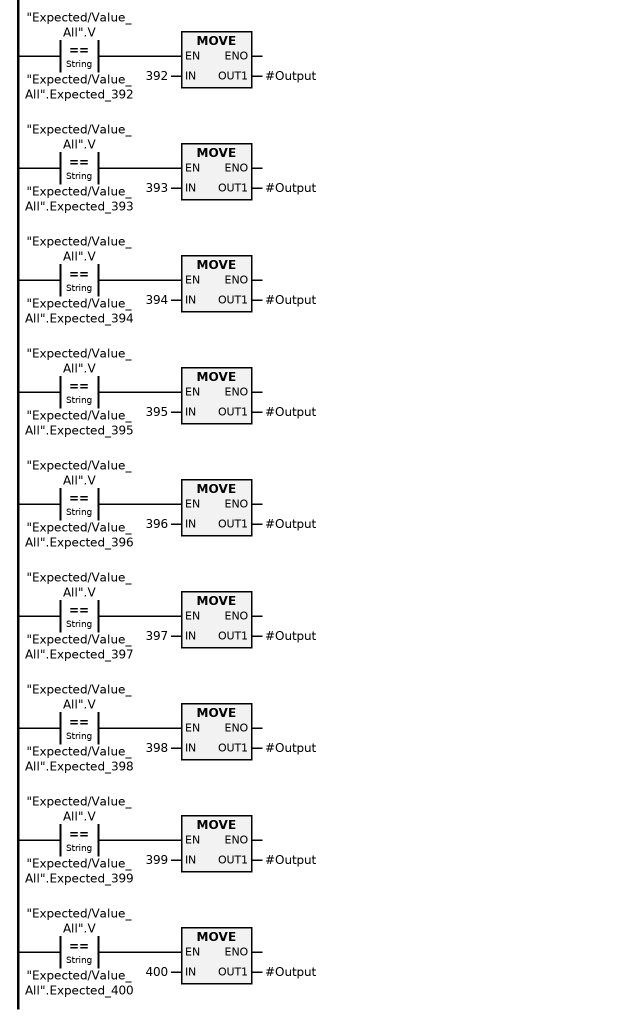
   RUNG wire#powerrail
      { S7_Templates := "SrcType := String" } EQ_Contact(in1 := "Expected/Value_All".V, in2 := "Expected/Value_All".Expected_381)
      Move(in := 381, out1 => #Output)
   END_RUNG
   RUNG wire#powerrail
      { S7_Templates := "SrcType := String" } EQ_Contact(in1 := "Expected/Value_All".V, in2 := "Expected/Value_All".Expected_382)
      Move(in := 382, out1 => #Output)
   END_RUNG
   RUNG wire#powerrail
      { S7_Templates := "SrcType := String" } EQ_Contact(in1 := "Expected/Value_All".V, in2 := "Expected/Value_All".Expected_383)
      Move(in := 383, out1 => #Output)
   END_RUNG
   RUNG wire#powerrail
      { S7_Templates := "SrcType := String" } EQ_Contact(in1 := "Expected/Value_All".V, in2 := "Expected/Value_All".Expected_384)
      Move(in := 384, out1 => #Output)
   END_RUNG
   RUNG wire#powerrail
      { S7_Templates := "SrcType := String" } EQ_Contact(in1 := "Expected/Value_All".V, in2 := "Expected/Value_All".Expected_385)
      Move(in := 385, out1 => #Output)
   END_RUNG
   RUNG wire#powerrail
      { S7_Templates := "SrcType := String" } EQ_Contact(in1 := "Expected/Value_All".V, in2 := "Expected/Value_All".Expected_386)
      Move(in := 386, out1 => #Output)
   END_RUNG
   RUNG wire#powerrail
      { S7_Templates := "SrcType := String" } EQ_Contact(in1 := "Expected/Value_All".V, in2 := "Expected/Value_All".Expected_387)
      Move(in := 387, out1 => #Output)
   END_RUNG
   RUNG wire#powerrail
      { S7_Templates := "SrcType := String" } EQ_Contact(in1 := "Expected/Value_All".V, in2 := "Expected/Value_All".Expected_388)
      Move(in := 388, out1 => #Output)
   END_RUNG
   RUNG wire#powerrail
      { S7_Templates := "SrcType := String" } EQ_Contact(in1 := "Expected/Value_All".V, in2 := "Expected/Value_All".Expected_389)
      Move(in := 389, out1 => #Output)
   END_RUNG
   RUNG wire#powerrail
      { S7_Templates := "SrcType := String" } EQ_Contact(in1 := "Expected/Value_All".V, in2 := "Expected/Value_All".Expected_390)
      Move(in := 390, out1 => #Output)
   END_RUNG
   RUNG wire#powerrail
      { S7_Templates := "SrcType := String" } EQ_Contact(in1 := "Expected/Value_All".V, in2 := "Expected/Value_All".Expected_391)
      Move(in := 391, out1 => #Output)
   END_RUNG
   RUNG wire#powerrail
      { S7_Templates := "SrcType := String" } EQ_Contact(in1 := "Expected/Value_All".V, in2 := "Expected/Value_All".Expected_392)
      Move(in := 392, out1 => #Output)
   END_RUNG
   RUNG wire#powerrail
      { S7_Templates := "SrcType := String" } EQ_Contact(in1 := "Expected/Value_All".V, in2 := "Expected/Value_All".Expected_393)
      Move(in := 393, out1 => #Output)
   END_RUNG
   RUNG wire#powerrail
      { S7_Templates := "SrcType := String" } EQ_Contact(in1 := "Expected/Value_All".V, in2 := "Expected/Value_All".Expected_394)
      Move(in := 394, out1 => #Output)
   END_RUNG
   RUNG wire#powerrail
      { S7_Templates := "SrcType := String" } EQ_Contact(in1 := "Expected/Value_All".V, in2 := "Expected/Value_All".Expected_395)
      Move(in := 395, out1 => #Output)
   END_RUNG
   RUNG wire#powerrail
      { S7_Templates := "SrcType := String" } EQ_Contact(in1 := "Expected/Value_All".V, in2 := "Expected/Value_All".Expected_396)
      Move(in := 396, out1 => #Output)
   END_RUNG
   RUNG wire#powerrail
      { S7_Templates := "SrcType := String" } EQ_Contact(in1 := "Expected/Value_All".V, in2 := "Expected/Value_All".Expected_397)
      Move(in := 397, out1 => #Output)
   END_RUNG
   RUNG wire#powerrail
      { S7_Templates := "SrcType := String" } EQ_Contact(in1 := "Expected/Value_All".V, in2 := "Expected/Value_All".Expected_398)
      Move(in := 398, out1 => #Output)
   END_RUNG
   RUNG wire#powerrail
      { S7_Templates := "SrcType := String" } EQ_Contact(in1 := "Expected/Value_All".V, in2 := "Expected/Value_All".Expected_399)
      Move(in := 399, out1 => #Output)
   END_RUNG
   RUNG wire#powerrail
      { S7_Templates := "SrcType := String" } EQ_Contact(in1 := "Expected/Value_All".V, in2 := "Expected/Value_All".Expected_400)
      Move(in := 400, out1 => #Output)
   END_RUNG
   // the same network as SCL:
   IF "Expected/Value_All".V = "Expected/Value_All".Expected_381 THEN #Output := 381; END_IF;
   IF "Expected/Value_All".V = "Expected/Value_All".Expected_382 THEN #Output := 382; END_IF;
   IF "Expected/Value_All".V = "Expected/Value_All".Expected_383 THEN #Output := 383; END_IF;
   IF "Expected/Value_All".V = "Expected/Value_All".Expected_384 THEN #Output := 384; END_IF;
   IF "Expected/Value_All".V = "Expected/Value_All".Expected_385 THEN #Output := 385; END_IF;
   IF "Expected/Value_All".V = "Expected/Value_All".Expected_386 THEN #Output := 386; END_IF;
   IF "Expected/Value_All".V = "Expected/Value_All".Expected_387 THEN #Output := 387; END_IF;
   IF "Expected/Value_All".V = "Expected/Value_All".Expected_388 THEN #Output := 388; END_IF;
   IF "Expected/Value_All".V = "Expected/Value_All".Expected_389 THEN #Output := 389; END_IF;
   IF "Expected/Value_All".V = "Expected/Value_All".Expected_390 THEN #Output := 390; END_IF;
   IF "Expected/Value_All".V = "Expected/Value_All".Expected_391 THEN #Output := 391; END_IF;
   IF "Expected/Value_All".V = "Expected/Value_All".Expected_392 THEN #Output := 392; END_IF;
   IF "Expected/Value_All".V = "Expected/Value_All".Expected_393 THEN #Output := 393; END_IF;
   IF "Expected/Value_All".V = "Expected/Value_All".Expected_394 THEN #Output := 394; END_IF;
   IF "Expected/Value_All".V = "Expected/Value_All".Expected_395 THEN #Output := 395; END_IF;
   IF "Expected/Value_All".V = "Expected/Value_All".Expected_396 THEN #Output := 396; END_IF;
   IF "Expected/Value_All".V = "Expected/Value_All".Expected_397 THEN #Output := 397; END_IF;
   IF "Expected/Value_All".V = "Expected/Value_All".Expected_398 THEN #Output := 398; END_IF;
   IF "Expected/Value_All".V = "Expected/Value_All".Expected_399 THEN #Output := 399; END_IF;
   IF "Expected/Value_All".V = "Expected/Value_All".Expected_400 THEN #Output := 400; END_IF;
END_REGION

REGION Network 21
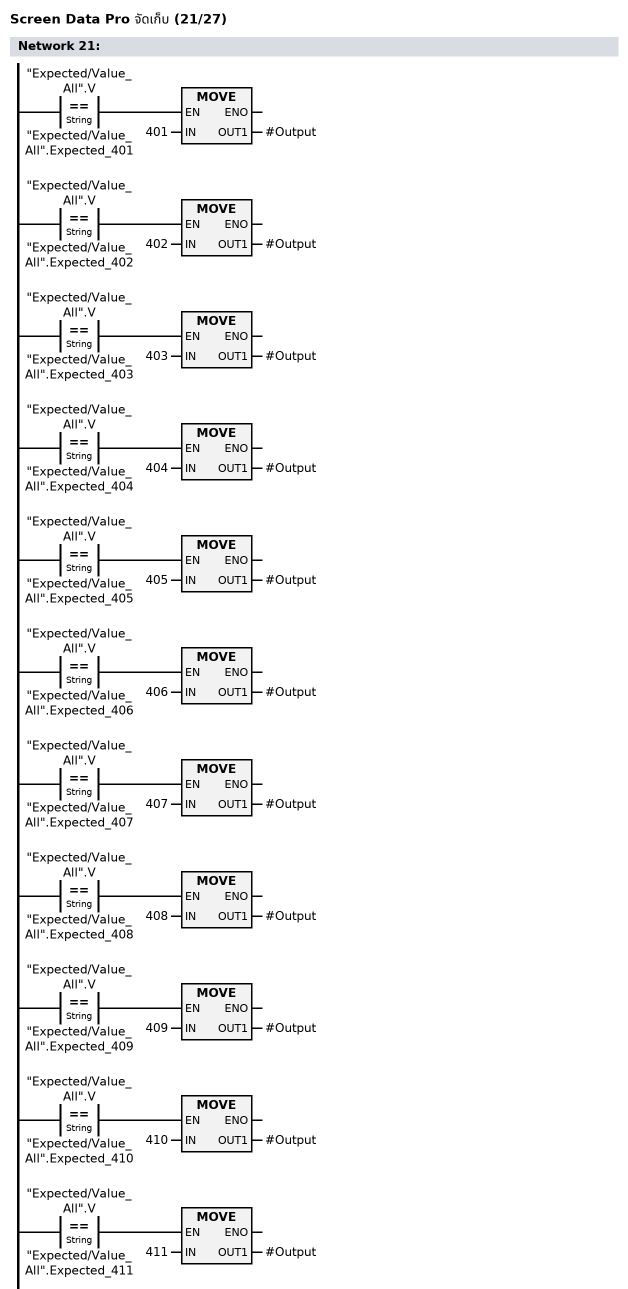
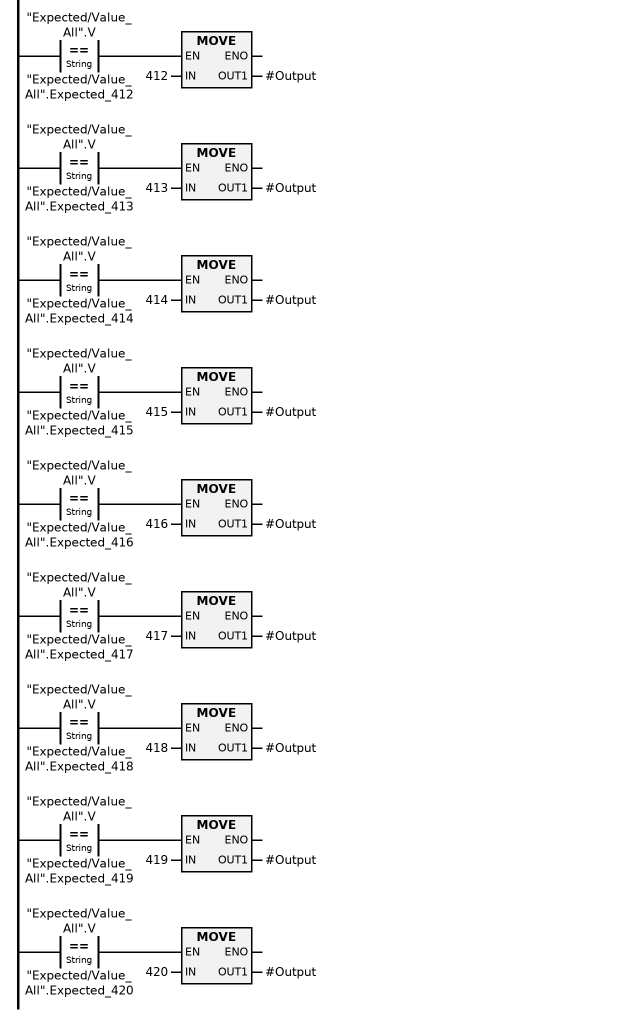
   RUNG wire#powerrail
      { S7_Templates := "SrcType := String" } EQ_Contact(in1 := "Expected/Value_All".V, in2 := "Expected/Value_All".Expected_401)
      Move(in := 401, out1 => #Output)
   END_RUNG
   RUNG wire#powerrail
      { S7_Templates := "SrcType := String" } EQ_Contact(in1 := "Expected/Value_All".V, in2 := "Expected/Value_All".Expected_402)
      Move(in := 402, out1 => #Output)
   END_RUNG
   RUNG wire#powerrail
      { S7_Templates := "SrcType := String" } EQ_Contact(in1 := "Expected/Value_All".V, in2 := "Expected/Value_All".Expected_403)
      Move(in := 403, out1 => #Output)
   END_RUNG
   RUNG wire#powerrail
      { S7_Templates := "SrcType := String" } EQ_Contact(in1 := "Expected/Value_All".V, in2 := "Expected/Value_All".Expected_404)
      Move(in := 404, out1 => #Output)
   END_RUNG
   RUNG wire#powerrail
      { S7_Templates := "SrcType := String" } EQ_Contact(in1 := "Expected/Value_All".V, in2 := "Expected/Value_All".Expected_405)
      Move(in := 405, out1 => #Output)
   END_RUNG
   RUNG wire#powerrail
      { S7_Templates := "SrcType := String" } EQ_Contact(in1 := "Expected/Value_All".V, in2 := "Expected/Value_All".Expected_406)
      Move(in := 406, out1 => #Output)
   END_RUNG
   RUNG wire#powerrail
      { S7_Templates := "SrcType := String" } EQ_Contact(in1 := "Expected/Value_All".V, in2 := "Expected/Value_All".Expected_407)
      Move(in := 407, out1 => #Output)
   END_RUNG
   RUNG wire#powerrail
      { S7_Templates := "SrcType := String" } EQ_Contact(in1 := "Expected/Value_All".V, in2 := "Expected/Value_All".Expected_408)
      Move(in := 408, out1 => #Output)
   END_RUNG
   RUNG wire#powerrail
      { S7_Templates := "SrcType := String" } EQ_Contact(in1 := "Expected/Value_All".V, in2 := "Expected/Value_All".Expected_409)
      Move(in := 409, out1 => #Output)
   END_RUNG
   RUNG wire#powerrail
      { S7_Templates := "SrcType := String" } EQ_Contact(in1 := "Expected/Value_All".V, in2 := "Expected/Value_All".Expected_410)
      Move(in := 410, out1 => #Output)
   END_RUNG
   RUNG wire#powerrail
      { S7_Templates := "SrcType := String" } EQ_Contact(in1 := "Expected/Value_All".V, in2 := "Expected/Value_All".Expected_411)
      Move(in := 411, out1 => #Output)
   END_RUNG
   RUNG wire#powerrail
      { S7_Templates := "SrcType := String" } EQ_Contact(in1 := "Expected/Value_All".V, in2 := "Expected/Value_All".Expected_412)
      Move(in := 412, out1 => #Output)
   END_RUNG
   RUNG wire#powerrail
      { S7_Templates := "SrcType := String" } EQ_Contact(in1 := "Expected/Value_All".V, in2 := "Expected/Value_All".Expected_413)
      Move(in := 413, out1 => #Output)
   END_RUNG
   RUNG wire#powerrail
      { S7_Templates := "SrcType := String" } EQ_Contact(in1 := "Expected/Value_All".V, in2 := "Expected/Value_All".Expected_414)
      Move(in := 414, out1 => #Output)
   END_RUNG
   RUNG wire#powerrail
      { S7_Templates := "SrcType := String" } EQ_Contact(in1 := "Expected/Value_All".V, in2 := "Expected/Value_All".Expected_415)
      Move(in := 415, out1 => #Output)
   END_RUNG
   RUNG wire#powerrail
      { S7_Templates := "SrcType := String" } EQ_Contact(in1 := "Expected/Value_All".V, in2 := "Expected/Value_All".Expected_416)
      Move(in := 416, out1 => #Output)
   END_RUNG
   RUNG wire#powerrail
      { S7_Templates := "SrcType := String" } EQ_Contact(in1 := "Expected/Value_All".V, in2 := "Expected/Value_All".Expected_417)
      Move(in := 417, out1 => #Output)
   END_RUNG
   RUNG wire#powerrail
      { S7_Templates := "SrcType := String" } EQ_Contact(in1 := "Expected/Value_All".V, in2 := "Expected/Value_All".Expected_418)
      Move(in := 418, out1 => #Output)
   END_RUNG
   RUNG wire#powerrail
      { S7_Templates := "SrcType := String" } EQ_Contact(in1 := "Expected/Value_All".V, in2 := "Expected/Value_All".Expected_419)
      Move(in := 419, out1 => #Output)
   END_RUNG
   RUNG wire#powerrail
      { S7_Templates := "SrcType := String" } EQ_Contact(in1 := "Expected/Value_All".V, in2 := "Expected/Value_All".Expected_420)
      Move(in := 420, out1 => #Output)
   END_RUNG
   // the same network as SCL:
   IF "Expected/Value_All".V = "Expected/Value_All".Expected_401 THEN #Output := 401; END_IF;
   IF "Expected/Value_All".V = "Expected/Value_All".Expected_402 THEN #Output := 402; END_IF;
   IF "Expected/Value_All".V = "Expected/Value_All".Expected_403 THEN #Output := 403; END_IF;
   IF "Expected/Value_All".V = "Expected/Value_All".Expected_404 THEN #Output := 404; END_IF;
   IF "Expected/Value_All".V = "Expected/Value_All".Expected_405 THEN #Output := 405; END_IF;
   IF "Expected/Value_All".V = "Expected/Value_All".Expected_406 THEN #Output := 406; END_IF;
   IF "Expected/Value_All".V = "Expected/Value_All".Expected_407 THEN #Output := 407; END_IF;
   IF "Expected/Value_All".V = "Expected/Value_All".Expected_408 THEN #Output := 408; END_IF;
   IF "Expected/Value_All".V = "Expected/Value_All".Expected_409 THEN #Output := 409; END_IF;
   IF "Expected/Value_All".V = "Expected/Value_All".Expected_410 THEN #Output := 410; END_IF;
   IF "Expected/Value_All".V = "Expected/Value_All".Expected_411 THEN #Output := 411; END_IF;
   IF "Expected/Value_All".V = "Expected/Value_All".Expected_412 THEN #Output := 412; END_IF;
   IF "Expected/Value_All".V = "Expected/Value_All".Expected_413 THEN #Output := 413; END_IF;
   IF "Expected/Value_All".V = "Expected/Value_All".Expected_414 THEN #Output := 414; END_IF;
   IF "Expected/Value_All".V = "Expected/Value_All".Expected_415 THEN #Output := 415; END_IF;
   IF "Expected/Value_All".V = "Expected/Value_All".Expected_416 THEN #Output := 416; END_IF;
   IF "Expected/Value_All".V = "Expected/Value_All".Expected_417 THEN #Output := 417; END_IF;
   IF "Expected/Value_All".V = "Expected/Value_All".Expected_418 THEN #Output := 418; END_IF;
   IF "Expected/Value_All".V = "Expected/Value_All".Expected_419 THEN #Output := 419; END_IF;
   IF "Expected/Value_All".V = "Expected/Value_All".Expected_420 THEN #Output := 420; END_IF;
END_REGION

REGION Network 22
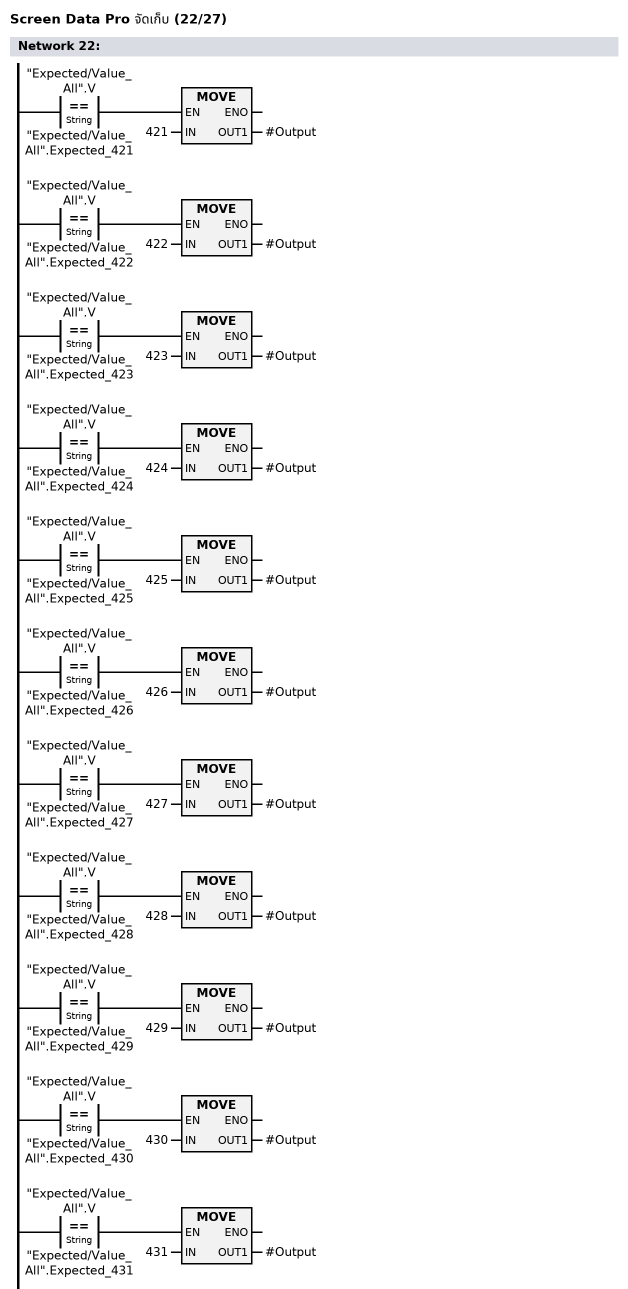
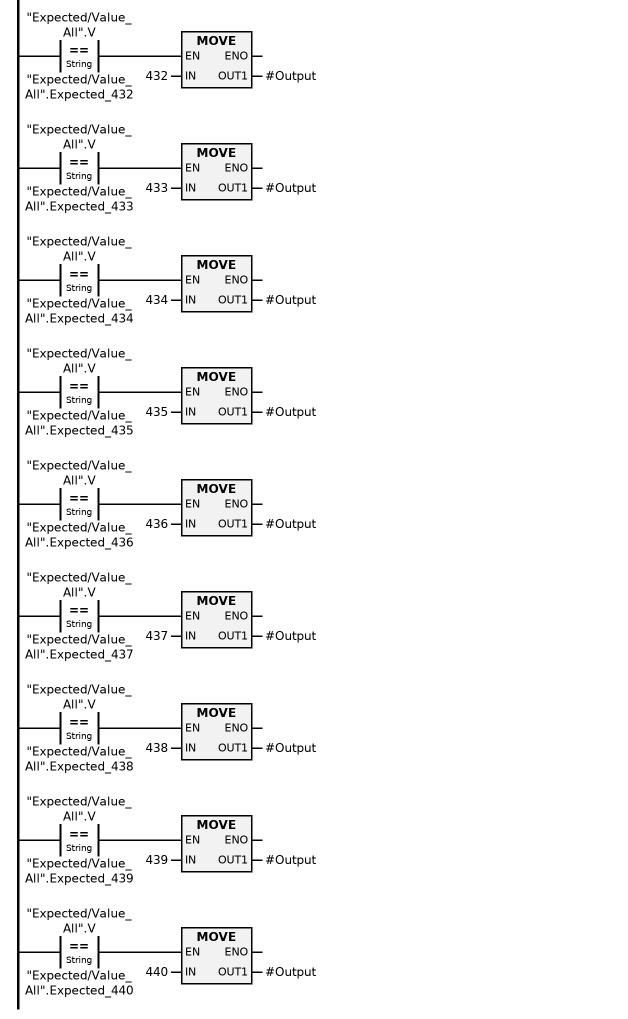
   RUNG wire#powerrail
      { S7_Templates := "SrcType := String" } EQ_Contact(in1 := "Expected/Value_All".V, in2 := "Expected/Value_All".Expected_421)
      Move(in := 421, out1 => #Output)
   END_RUNG
   RUNG wire#powerrail
      { S7_Templates := "SrcType := String" } EQ_Contact(in1 := "Expected/Value_All".V, in2 := "Expected/Value_All".Expected_422)
      Move(in := 422, out1 => #Output)
   END_RUNG
   RUNG wire#powerrail
      { S7_Templates := "SrcType := String" } EQ_Contact(in1 := "Expected/Value_All".V, in2 := "Expected/Value_All".Expected_423)
      Move(in := 423, out1 => #Output)
   END_RUNG
   RUNG wire#powerrail
      { S7_Templates := "SrcType := String" } EQ_Contact(in1 := "Expected/Value_All".V, in2 := "Expected/Value_All".Expected_424)
      Move(in := 424, out1 => #Output)
   END_RUNG
   RUNG wire#powerrail
      { S7_Templates := "SrcType := String" } EQ_Contact(in1 := "Expected/Value_All".V, in2 := "Expected/Value_All".Expected_425)
      Move(in := 425, out1 => #Output)
   END_RUNG
   RUNG wire#powerrail
      { S7_Templates := "SrcType := String" } EQ_Contact(in1 := "Expected/Value_All".V, in2 := "Expected/Value_All".Expected_426)
      Move(in := 426, out1 => #Output)
   END_RUNG
   RUNG wire#powerrail
      { S7_Templates := "SrcType := String" } EQ_Contact(in1 := "Expected/Value_All".V, in2 := "Expected/Value_All".Expected_427)
      Move(in := 427, out1 => #Output)
   END_RUNG
   RUNG wire#powerrail
      { S7_Templates := "SrcType := String" } EQ_Contact(in1 := "Expected/Value_All".V, in2 := "Expected/Value_All".Expected_428)
      Move(in := 428, out1 => #Output)
   END_RUNG
   RUNG wire#powerrail
      { S7_Templates := "SrcType := String" } EQ_Contact(in1 := "Expected/Value_All".V, in2 := "Expected/Value_All".Expected_429)
      Move(in := 429, out1 => #Output)
   END_RUNG
   RUNG wire#powerrail
      { S7_Templates := "SrcType := String" } EQ_Contact(in1 := "Expected/Value_All".V, in2 := "Expected/Value_All".Expected_430)
      Move(in := 430, out1 => #Output)
   END_RUNG
   RUNG wire#powerrail
      { S7_Templates := "SrcType := String" } EQ_Contact(in1 := "Expected/Value_All".V, in2 := "Expected/Value_All".Expected_431)
      Move(in := 431, out1 => #Output)
   END_RUNG
   RUNG wire#powerrail
      { S7_Templates := "SrcType := String" } EQ_Contact(in1 := "Expected/Value_All".V, in2 := "Expected/Value_All".Expected_432)
      Move(in := 432, out1 => #Output)
   END_RUNG
   RUNG wire#powerrail
      { S7_Templates := "SrcType := String" } EQ_Contact(in1 := "Expected/Value_All".V, in2 := "Expected/Value_All".Expected_433)
      Move(in := 433, out1 => #Output)
   END_RUNG
   RUNG wire#powerrail
      { S7_Templates := "SrcType := String" } EQ_Contact(in1 := "Expected/Value_All".V, in2 := "Expected/Value_All".Expected_434)
      Move(in := 434, out1 => #Output)
   END_RUNG
   RUNG wire#powerrail
      { S7_Templates := "SrcType := String" } EQ_Contact(in1 := "Expected/Value_All".V, in2 := "Expected/Value_All".Expected_435)
      Move(in := 435, out1 => #Output)
   END_RUNG
   RUNG wire#powerrail
      { S7_Templates := "SrcType := String" } EQ_Contact(in1 := "Expected/Value_All".V, in2 := "Expected/Value_All".Expected_436)
      Move(in := 436, out1 => #Output)
   END_RUNG
   RUNG wire#powerrail
      { S7_Templates := "SrcType := String" } EQ_Contact(in1 := "Expected/Value_All".V, in2 := "Expected/Value_All".Expected_437)
      Move(in := 437, out1 => #Output)
   END_RUNG
   RUNG wire#powerrail
      { S7_Templates := "SrcType := String" } EQ_Contact(in1 := "Expected/Value_All".V, in2 := "Expected/Value_All".Expected_438)
      Move(in := 438, out1 => #Output)
   END_RUNG
   RUNG wire#powerrail
      { S7_Templates := "SrcType := String" } EQ_Contact(in1 := "Expected/Value_All".V, in2 := "Expected/Value_All".Expected_439)
      Move(in := 439, out1 => #Output)
   END_RUNG
   RUNG wire#powerrail
      { S7_Templates := "SrcType := String" } EQ_Contact(in1 := "Expected/Value_All".V, in2 := "Expected/Value_All".Expected_440)
      Move(in := 440, out1 => #Output)
   END_RUNG
   // the same network as SCL:
   IF "Expected/Value_All".V = "Expected/Value_All".Expected_421 THEN #Output := 421; END_IF;
   IF "Expected/Value_All".V = "Expected/Value_All".Expected_422 THEN #Output := 422; END_IF;
   IF "Expected/Value_All".V = "Expected/Value_All".Expected_423 THEN #Output := 423; END_IF;
   IF "Expected/Value_All".V = "Expected/Value_All".Expected_424 THEN #Output := 424; END_IF;
   IF "Expected/Value_All".V = "Expected/Value_All".Expected_425 THEN #Output := 425; END_IF;
   IF "Expected/Value_All".V = "Expected/Value_All".Expected_426 THEN #Output := 426; END_IF;
   IF "Expected/Value_All".V = "Expected/Value_All".Expected_427 THEN #Output := 427; END_IF;
   IF "Expected/Value_All".V = "Expected/Value_All".Expected_428 THEN #Output := 428; END_IF;
   IF "Expected/Value_All".V = "Expected/Value_All".Expected_429 THEN #Output := 429; END_IF;
   IF "Expected/Value_All".V = "Expected/Value_All".Expected_430 THEN #Output := 430; END_IF;
   IF "Expected/Value_All".V = "Expected/Value_All".Expected_431 THEN #Output := 431; END_IF;
   IF "Expected/Value_All".V = "Expected/Value_All".Expected_432 THEN #Output := 432; END_IF;
   IF "Expected/Value_All".V = "Expected/Value_All".Expected_433 THEN #Output := 433; END_IF;
   IF "Expected/Value_All".V = "Expected/Value_All".Expected_434 THEN #Output := 434; END_IF;
   IF "Expected/Value_All".V = "Expected/Value_All".Expected_435 THEN #Output := 435; END_IF;
   IF "Expected/Value_All".V = "Expected/Value_All".Expected_436 THEN #Output := 436; END_IF;
   IF "Expected/Value_All".V = "Expected/Value_All".Expected_437 THEN #Output := 437; END_IF;
   IF "Expected/Value_All".V = "Expected/Value_All".Expected_438 THEN #Output := 438; END_IF;
   IF "Expected/Value_All".V = "Expected/Value_All".Expected_439 THEN #Output := 439; END_IF;
   IF "Expected/Value_All".V = "Expected/Value_All".Expected_440 THEN #Output := 440; END_IF;
END_REGION

REGION Network 23
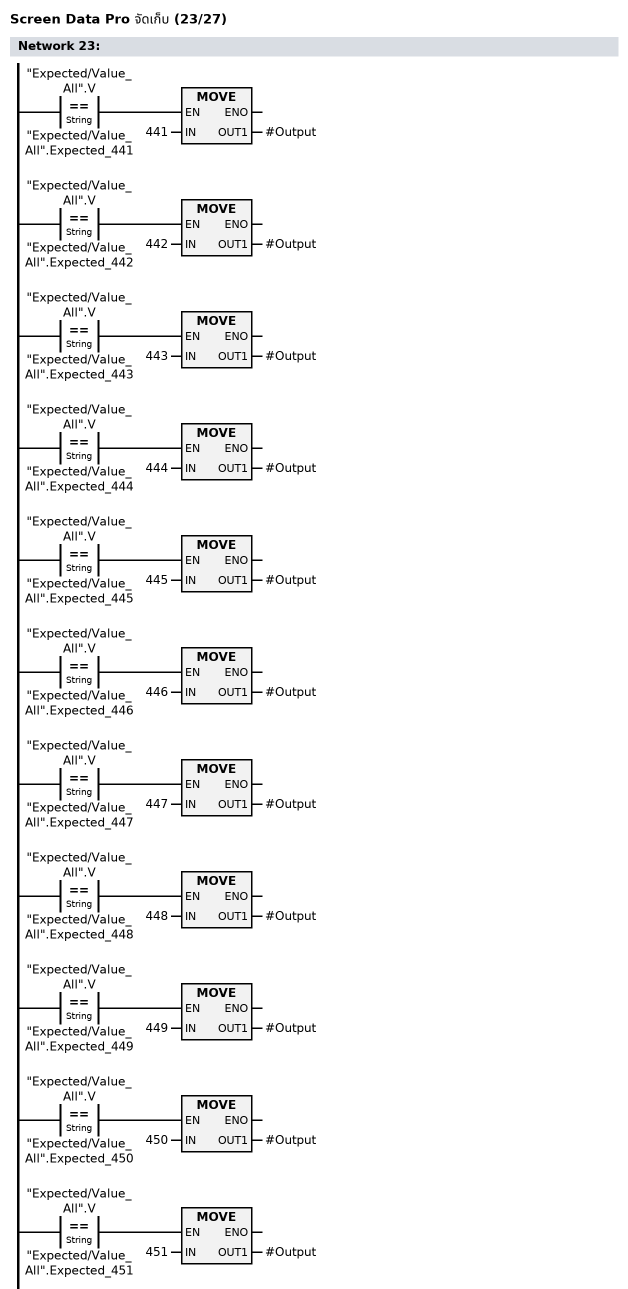
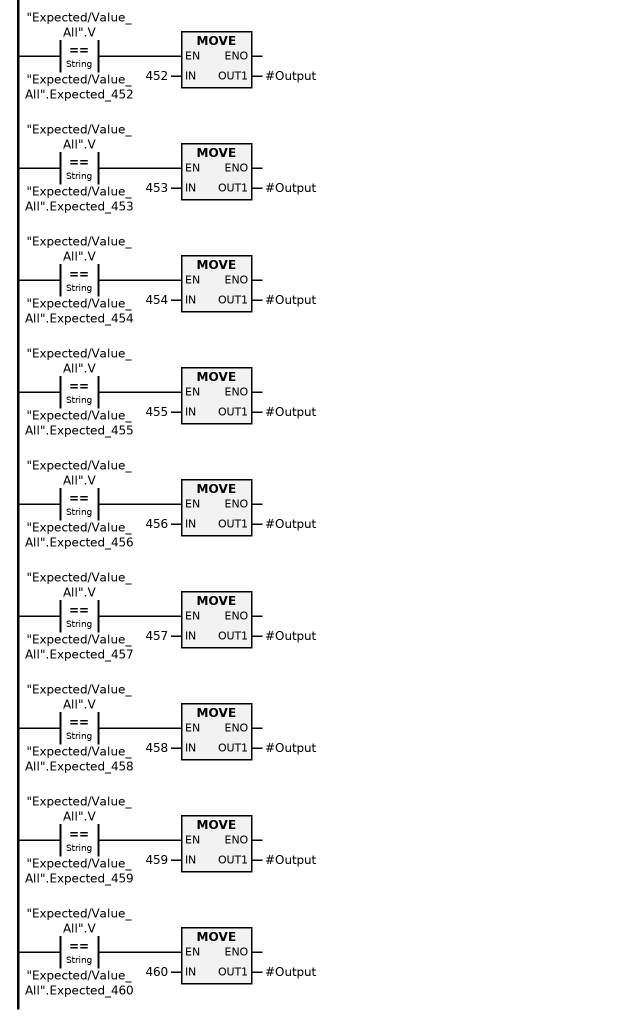
   RUNG wire#powerrail
      { S7_Templates := "SrcType := String" } EQ_Contact(in1 := "Expected/Value_All".V, in2 := "Expected/Value_All".Expected_441)
      Move(in := 441, out1 => #Output)
   END_RUNG
   RUNG wire#powerrail
      { S7_Templates := "SrcType := String" } EQ_Contact(in1 := "Expected/Value_All".V, in2 := "Expected/Value_All".Expected_442)
      Move(in := 442, out1 => #Output)
   END_RUNG
   RUNG wire#powerrail
      { S7_Templates := "SrcType := String" } EQ_Contact(in1 := "Expected/Value_All".V, in2 := "Expected/Value_All".Expected_443)
      Move(in := 443, out1 => #Output)
   END_RUNG
   RUNG wire#powerrail
      { S7_Templates := "SrcType := String" } EQ_Contact(in1 := "Expected/Value_All".V, in2 := "Expected/Value_All".Expected_444)
      Move(in := 444, out1 => #Output)
   END_RUNG
   RUNG wire#powerrail
      { S7_Templates := "SrcType := String" } EQ_Contact(in1 := "Expected/Value_All".V, in2 := "Expected/Value_All".Expected_445)
      Move(in := 445, out1 => #Output)
   END_RUNG
   RUNG wire#powerrail
      { S7_Templates := "SrcType := String" } EQ_Contact(in1 := "Expected/Value_All".V, in2 := "Expected/Value_All".Expected_446)
      Move(in := 446, out1 => #Output)
   END_RUNG
   RUNG wire#powerrail
      { S7_Templates := "SrcType := String" } EQ_Contact(in1 := "Expected/Value_All".V, in2 := "Expected/Value_All".Expected_447)
      Move(in := 447, out1 => #Output)
   END_RUNG
   RUNG wire#powerrail
      { S7_Templates := "SrcType := String" } EQ_Contact(in1 := "Expected/Value_All".V, in2 := "Expected/Value_All".Expected_448)
      Move(in := 448, out1 => #Output)
   END_RUNG
   RUNG wire#powerrail
      { S7_Templates := "SrcType := String" } EQ_Contact(in1 := "Expected/Value_All".V, in2 := "Expected/Value_All".Expected_449)
      Move(in := 449, out1 => #Output)
   END_RUNG
   RUNG wire#powerrail
      { S7_Templates := "SrcType := String" } EQ_Contact(in1 := "Expected/Value_All".V, in2 := "Expected/Value_All".Expected_450)
      Move(in := 450, out1 => #Output)
   END_RUNG
   RUNG wire#powerrail
      { S7_Templates := "SrcType := String" } EQ_Contact(in1 := "Expected/Value_All".V, in2 := "Expected/Value_All".Expected_451)
      Move(in := 451, out1 => #Output)
   END_RUNG
   RUNG wire#powerrail
      { S7_Templates := "SrcType := String" } EQ_Contact(in1 := "Expected/Value_All".V, in2 := "Expected/Value_All".Expected_452)
      Move(in := 452, out1 => #Output)
   END_RUNG
   RUNG wire#powerrail
      { S7_Templates := "SrcType := String" } EQ_Contact(in1 := "Expected/Value_All".V, in2 := "Expected/Value_All".Expected_453)
      Move(in := 453, out1 => #Output)
   END_RUNG
   RUNG wire#powerrail
      { S7_Templates := "SrcType := String" } EQ_Contact(in1 := "Expected/Value_All".V, in2 := "Expected/Value_All".Expected_454)
      Move(in := 454, out1 => #Output)
   END_RUNG
   RUNG wire#powerrail
      { S7_Templates := "SrcType := String" } EQ_Contact(in1 := "Expected/Value_All".V, in2 := "Expected/Value_All".Expected_455)
      Move(in := 455, out1 => #Output)
   END_RUNG
   RUNG wire#powerrail
      { S7_Templates := "SrcType := String" } EQ_Contact(in1 := "Expected/Value_All".V, in2 := "Expected/Value_All".Expected_456)
      Move(in := 456, out1 => #Output)
   END_RUNG
   RUNG wire#powerrail
      { S7_Templates := "SrcType := String" } EQ_Contact(in1 := "Expected/Value_All".V, in2 := "Expected/Value_All".Expected_457)
      Move(in := 457, out1 => #Output)
   END_RUNG
   RUNG wire#powerrail
      { S7_Templates := "SrcType := String" } EQ_Contact(in1 := "Expected/Value_All".V, in2 := "Expected/Value_All".Expected_458)
      Move(in := 458, out1 => #Output)
   END_RUNG
   RUNG wire#powerrail
      { S7_Templates := "SrcType := String" } EQ_Contact(in1 := "Expected/Value_All".V, in2 := "Expected/Value_All".Expected_459)
      Move(in := 459, out1 => #Output)
   END_RUNG
   RUNG wire#powerrail
      { S7_Templates := "SrcType := String" } EQ_Contact(in1 := "Expected/Value_All".V, in2 := "Expected/Value_All".Expected_460)
      Move(in := 460, out1 => #Output)
   END_RUNG
   // the same network as SCL:
   IF "Expected/Value_All".V = "Expected/Value_All".Expected_441 THEN #Output := 441; END_IF;
   IF "Expected/Value_All".V = "Expected/Value_All".Expected_442 THEN #Output := 442; END_IF;
   IF "Expected/Value_All".V = "Expected/Value_All".Expected_443 THEN #Output := 443; END_IF;
   IF "Expected/Value_All".V = "Expected/Value_All".Expected_444 THEN #Output := 444; END_IF;
   IF "Expected/Value_All".V = "Expected/Value_All".Expected_445 THEN #Output := 445; END_IF;
   IF "Expected/Value_All".V = "Expected/Value_All".Expected_446 THEN #Output := 446; END_IF;
   IF "Expected/Value_All".V = "Expected/Value_All".Expected_447 THEN #Output := 447; END_IF;
   IF "Expected/Value_All".V = "Expected/Value_All".Expected_448 THEN #Output := 448; END_IF;
   IF "Expected/Value_All".V = "Expected/Value_All".Expected_449 THEN #Output := 449; END_IF;
   IF "Expected/Value_All".V = "Expected/Value_All".Expected_450 THEN #Output := 450; END_IF;
   IF "Expected/Value_All".V = "Expected/Value_All".Expected_451 THEN #Output := 451; END_IF;
   IF "Expected/Value_All".V = "Expected/Value_All".Expected_452 THEN #Output := 452; END_IF;
   IF "Expected/Value_All".V = "Expected/Value_All".Expected_453 THEN #Output := 453; END_IF;
   IF "Expected/Value_All".V = "Expected/Value_All".Expected_454 THEN #Output := 454; END_IF;
   IF "Expected/Value_All".V = "Expected/Value_All".Expected_455 THEN #Output := 455; END_IF;
   IF "Expected/Value_All".V = "Expected/Value_All".Expected_456 THEN #Output := 456; END_IF;
   IF "Expected/Value_All".V = "Expected/Value_All".Expected_457 THEN #Output := 457; END_IF;
   IF "Expected/Value_All".V = "Expected/Value_All".Expected_458 THEN #Output := 458; END_IF;
   IF "Expected/Value_All".V = "Expected/Value_All".Expected_459 THEN #Output := 459; END_IF;
   IF "Expected/Value_All".V = "Expected/Value_All".Expected_460 THEN #Output := 460; END_IF;
END_REGION

REGION Network 24
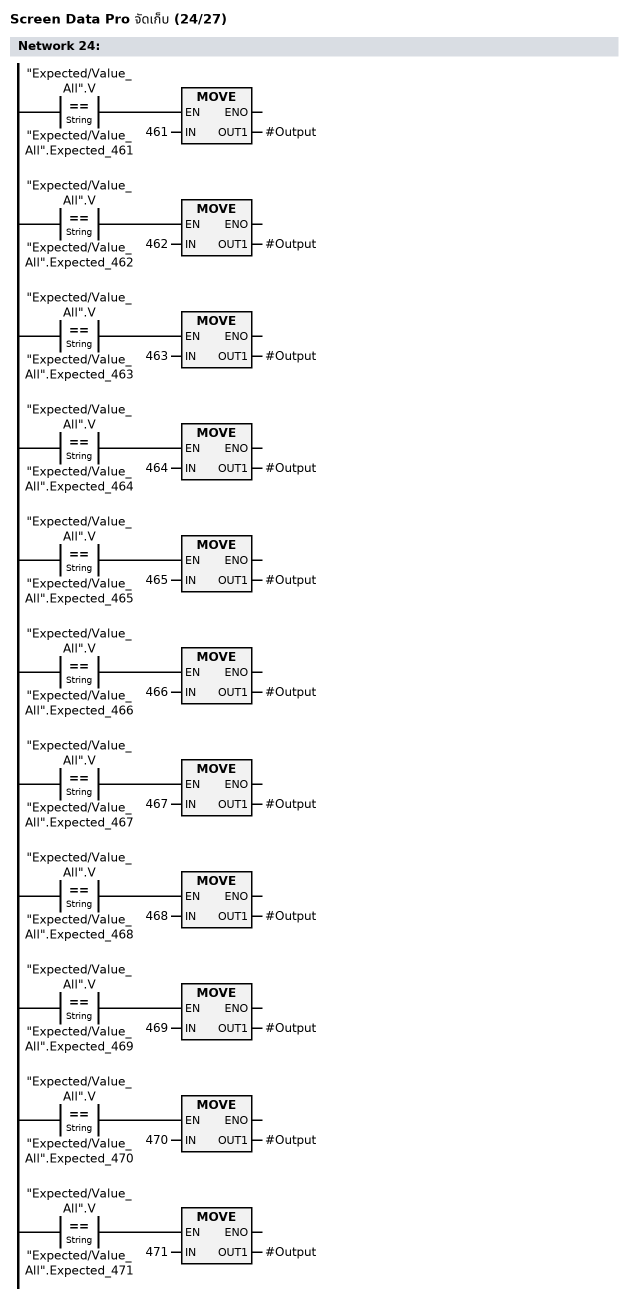
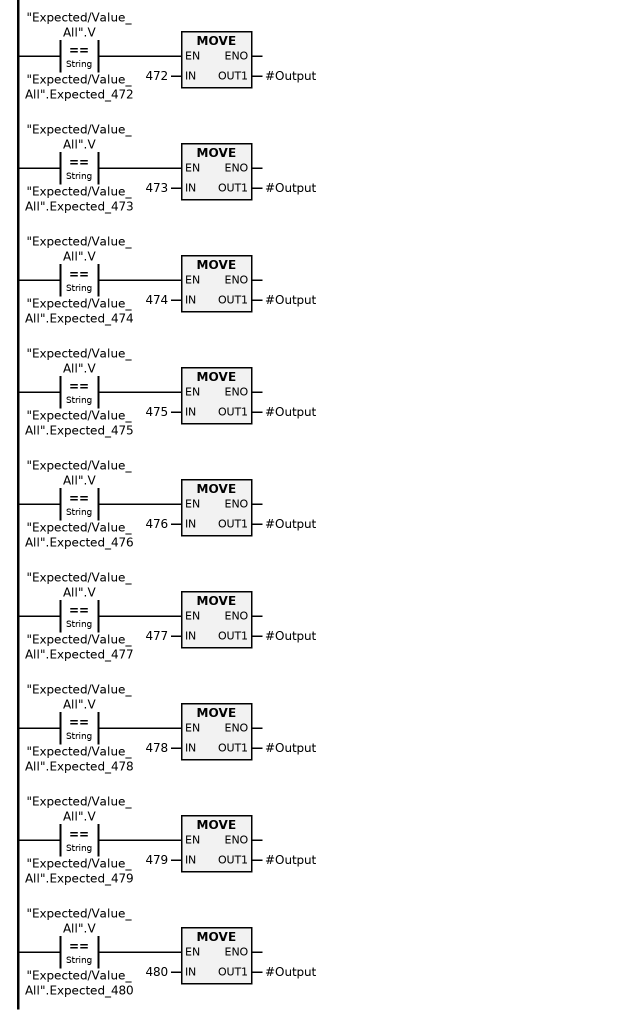
   RUNG wire#powerrail
      { S7_Templates := "SrcType := String" } EQ_Contact(in1 := "Expected/Value_All".V, in2 := "Expected/Value_All".Expected_461)
      Move(in := 461, out1 => #Output)
   END_RUNG
   RUNG wire#powerrail
      { S7_Templates := "SrcType := String" } EQ_Contact(in1 := "Expected/Value_All".V, in2 := "Expected/Value_All".Expected_462)
      Move(in := 462, out1 => #Output)
   END_RUNG
   RUNG wire#powerrail
      { S7_Templates := "SrcType := String" } EQ_Contact(in1 := "Expected/Value_All".V, in2 := "Expected/Value_All".Expected_463)
      Move(in := 463, out1 => #Output)
   END_RUNG
   RUNG wire#powerrail
      { S7_Templates := "SrcType := String" } EQ_Contact(in1 := "Expected/Value_All".V, in2 := "Expected/Value_All".Expected_464)
      Move(in := 464, out1 => #Output)
   END_RUNG
   RUNG wire#powerrail
      { S7_Templates := "SrcType := String" } EQ_Contact(in1 := "Expected/Value_All".V, in2 := "Expected/Value_All".Expected_465)
      Move(in := 465, out1 => #Output)
   END_RUNG
   RUNG wire#powerrail
      { S7_Templates := "SrcType := String" } EQ_Contact(in1 := "Expected/Value_All".V, in2 := "Expected/Value_All".Expected_466)
      Move(in := 466, out1 => #Output)
   END_RUNG
   RUNG wire#powerrail
      { S7_Templates := "SrcType := String" } EQ_Contact(in1 := "Expected/Value_All".V, in2 := "Expected/Value_All".Expected_467)
      Move(in := 467, out1 => #Output)
   END_RUNG
   RUNG wire#powerrail
      { S7_Templates := "SrcType := String" } EQ_Contact(in1 := "Expected/Value_All".V, in2 := "Expected/Value_All".Expected_468)
      Move(in := 468, out1 => #Output)
   END_RUNG
   RUNG wire#powerrail
      { S7_Templates := "SrcType := String" } EQ_Contact(in1 := "Expected/Value_All".V, in2 := "Expected/Value_All".Expected_469)
      Move(in := 469, out1 => #Output)
   END_RUNG
   RUNG wire#powerrail
      { S7_Templates := "SrcType := String" } EQ_Contact(in1 := "Expected/Value_All".V, in2 := "Expected/Value_All".Expected_470)
      Move(in := 470, out1 => #Output)
   END_RUNG
   RUNG wire#powerrail
      { S7_Templates := "SrcType := String" } EQ_Contact(in1 := "Expected/Value_All".V, in2 := "Expected/Value_All".Expected_471)
      Move(in := 471, out1 => #Output)
   END_RUNG
   RUNG wire#powerrail
      { S7_Templates := "SrcType := String" } EQ_Contact(in1 := "Expected/Value_All".V, in2 := "Expected/Value_All".Expected_472)
      Move(in := 472, out1 => #Output)
   END_RUNG
   RUNG wire#powerrail
      { S7_Templates := "SrcType := String" } EQ_Contact(in1 := "Expected/Value_All".V, in2 := "Expected/Value_All".Expected_473)
      Move(in := 473, out1 => #Output)
   END_RUNG
   RUNG wire#powerrail
      { S7_Templates := "SrcType := String" } EQ_Contact(in1 := "Expected/Value_All".V, in2 := "Expected/Value_All".Expected_474)
      Move(in := 474, out1 => #Output)
   END_RUNG
   RUNG wire#powerrail
      { S7_Templates := "SrcType := String" } EQ_Contact(in1 := "Expected/Value_All".V, in2 := "Expected/Value_All".Expected_475)
      Move(in := 475, out1 => #Output)
   END_RUNG
   RUNG wire#powerrail
      { S7_Templates := "SrcType := String" } EQ_Contact(in1 := "Expected/Value_All".V, in2 := "Expected/Value_All".Expected_476)
      Move(in := 476, out1 => #Output)
   END_RUNG
   RUNG wire#powerrail
      { S7_Templates := "SrcType := String" } EQ_Contact(in1 := "Expected/Value_All".V, in2 := "Expected/Value_All".Expected_477)
      Move(in := 477, out1 => #Output)
   END_RUNG
   RUNG wire#powerrail
      { S7_Templates := "SrcType := String" } EQ_Contact(in1 := "Expected/Value_All".V, in2 := "Expected/Value_All".Expected_478)
      Move(in := 478, out1 => #Output)
   END_RUNG
   RUNG wire#powerrail
      { S7_Templates := "SrcType := String" } EQ_Contact(in1 := "Expected/Value_All".V, in2 := "Expected/Value_All".Expected_479)
      Move(in := 479, out1 => #Output)
   END_RUNG
   RUNG wire#powerrail
      { S7_Templates := "SrcType := String" } EQ_Contact(in1 := "Expected/Value_All".V, in2 := "Expected/Value_All".Expected_480)
      Move(in := 480, out1 => #Output)
   END_RUNG
   // the same network as SCL:
   IF "Expected/Value_All".V = "Expected/Value_All".Expected_461 THEN #Output := 461; END_IF;
   IF "Expected/Value_All".V = "Expected/Value_All".Expected_462 THEN #Output := 462; END_IF;
   IF "Expected/Value_All".V = "Expected/Value_All".Expected_463 THEN #Output := 463; END_IF;
   IF "Expected/Value_All".V = "Expected/Value_All".Expected_464 THEN #Output := 464; END_IF;
   IF "Expected/Value_All".V = "Expected/Value_All".Expected_465 THEN #Output := 465; END_IF;
   IF "Expected/Value_All".V = "Expected/Value_All".Expected_466 THEN #Output := 466; END_IF;
   IF "Expected/Value_All".V = "Expected/Value_All".Expected_467 THEN #Output := 467; END_IF;
   IF "Expected/Value_All".V = "Expected/Value_All".Expected_468 THEN #Output := 468; END_IF;
   IF "Expected/Value_All".V = "Expected/Value_All".Expected_469 THEN #Output := 469; END_IF;
   IF "Expected/Value_All".V = "Expected/Value_All".Expected_470 THEN #Output := 470; END_IF;
   IF "Expected/Value_All".V = "Expected/Value_All".Expected_471 THEN #Output := 471; END_IF;
   IF "Expected/Value_All".V = "Expected/Value_All".Expected_472 THEN #Output := 472; END_IF;
   IF "Expected/Value_All".V = "Expected/Value_All".Expected_473 THEN #Output := 473; END_IF;
   IF "Expected/Value_All".V = "Expected/Value_All".Expected_474 THEN #Output := 474; END_IF;
   IF "Expected/Value_All".V = "Expected/Value_All".Expected_475 THEN #Output := 475; END_IF;
   IF "Expected/Value_All".V = "Expected/Value_All".Expected_476 THEN #Output := 476; END_IF;
   IF "Expected/Value_All".V = "Expected/Value_All".Expected_477 THEN #Output := 477; END_IF;
   IF "Expected/Value_All".V = "Expected/Value_All".Expected_478 THEN #Output := 478; END_IF;
   IF "Expected/Value_All".V = "Expected/Value_All".Expected_479 THEN #Output := 479; END_IF;
   IF "Expected/Value_All".V = "Expected/Value_All".Expected_480 THEN #Output := 480; END_IF;
END_REGION

REGION Network 25
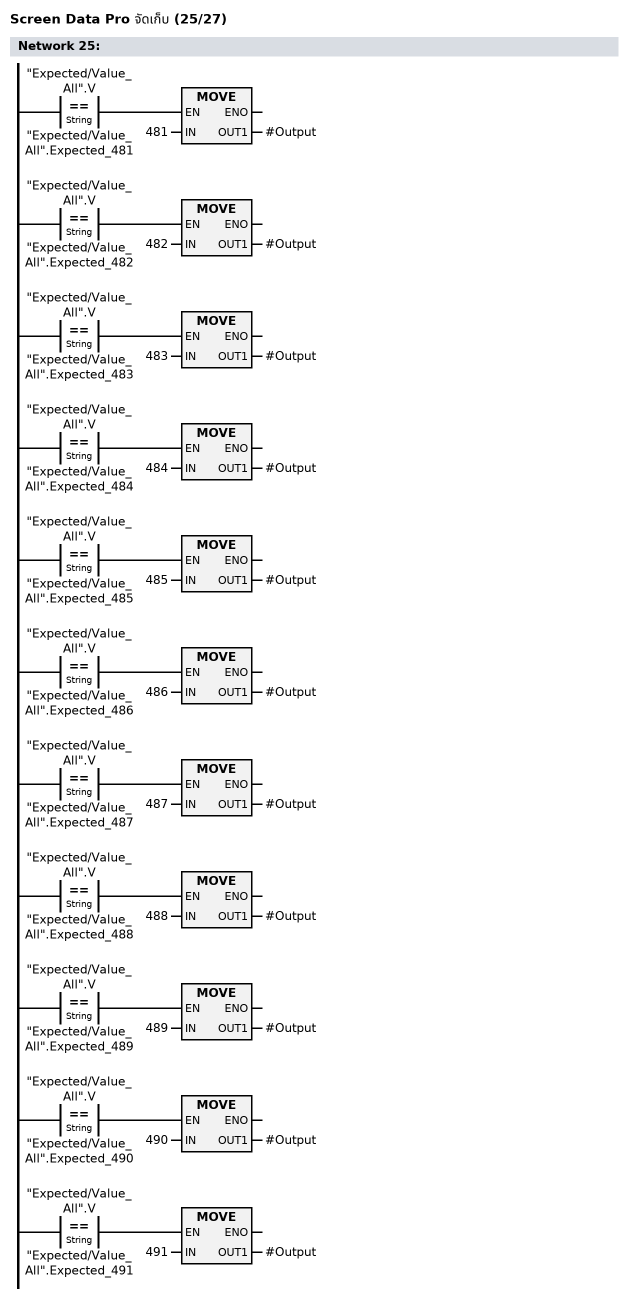
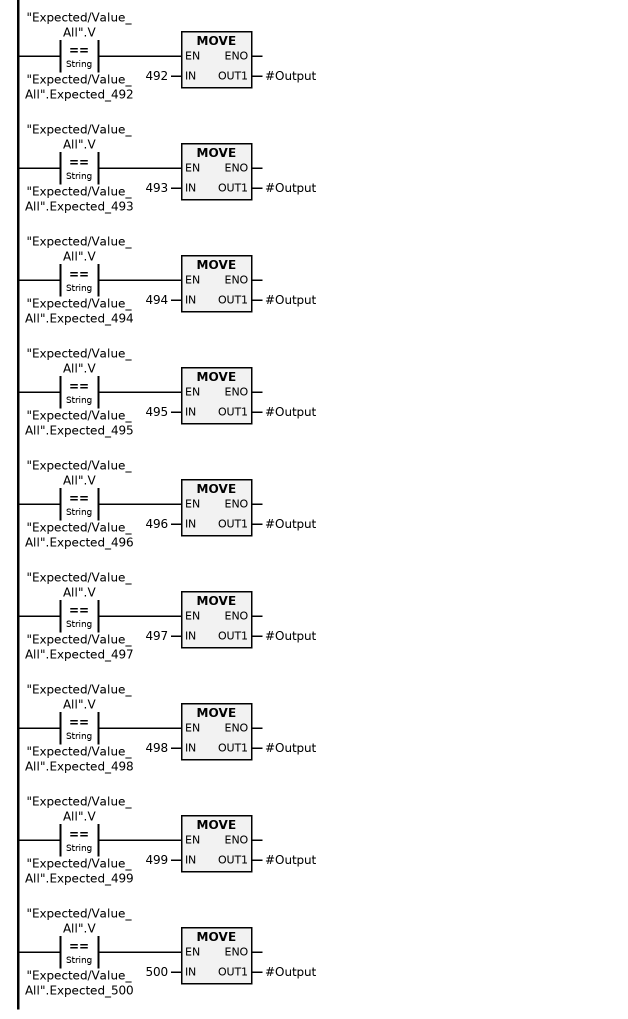
   RUNG wire#powerrail
      { S7_Templates := "SrcType := String" } EQ_Contact(in1 := "Expected/Value_All".V, in2 := "Expected/Value_All".Expected_481)
      Move(in := 481, out1 => #Output)
   END_RUNG
   RUNG wire#powerrail
      { S7_Templates := "SrcType := String" } EQ_Contact(in1 := "Expected/Value_All".V, in2 := "Expected/Value_All".Expected_482)
      Move(in := 482, out1 => #Output)
   END_RUNG
   RUNG wire#powerrail
      { S7_Templates := "SrcType := String" } EQ_Contact(in1 := "Expected/Value_All".V, in2 := "Expected/Value_All".Expected_483)
      Move(in := 483, out1 => #Output)
   END_RUNG
   RUNG wire#powerrail
      { S7_Templates := "SrcType := String" } EQ_Contact(in1 := "Expected/Value_All".V, in2 := "Expected/Value_All".Expected_484)
      Move(in := 484, out1 => #Output)
   END_RUNG
   RUNG wire#powerrail
      { S7_Templates := "SrcType := String" } EQ_Contact(in1 := "Expected/Value_All".V, in2 := "Expected/Value_All".Expected_485)
      Move(in := 485, out1 => #Output)
   END_RUNG
   RUNG wire#powerrail
      { S7_Templates := "SrcType := String" } EQ_Contact(in1 := "Expected/Value_All".V, in2 := "Expected/Value_All".Expected_486)
      Move(in := 486, out1 => #Output)
   END_RUNG
   RUNG wire#powerrail
      { S7_Templates := "SrcType := String" } EQ_Contact(in1 := "Expected/Value_All".V, in2 := "Expected/Value_All".Expected_487)
      Move(in := 487, out1 => #Output)
   END_RUNG
   RUNG wire#powerrail
      { S7_Templates := "SrcType := String" } EQ_Contact(in1 := "Expected/Value_All".V, in2 := "Expected/Value_All".Expected_488)
      Move(in := 488, out1 => #Output)
   END_RUNG
   RUNG wire#powerrail
      { S7_Templates := "SrcType := String" } EQ_Contact(in1 := "Expected/Value_All".V, in2 := "Expected/Value_All".Expected_489)
      Move(in := 489, out1 => #Output)
   END_RUNG
   RUNG wire#powerrail
      { S7_Templates := "SrcType := String" } EQ_Contact(in1 := "Expected/Value_All".V, in2 := "Expected/Value_All".Expected_490)
      Move(in := 490, out1 => #Output)
   END_RUNG
   RUNG wire#powerrail
      { S7_Templates := "SrcType := String" } EQ_Contact(in1 := "Expected/Value_All".V, in2 := "Expected/Value_All".Expected_491)
      Move(in := 491, out1 => #Output)
   END_RUNG
   RUNG wire#powerrail
      { S7_Templates := "SrcType := String" } EQ_Contact(in1 := "Expected/Value_All".V, in2 := "Expected/Value_All".Expected_492)
      Move(in := 492, out1 => #Output)
   END_RUNG
   RUNG wire#powerrail
      { S7_Templates := "SrcType := String" } EQ_Contact(in1 := "Expected/Value_All".V, in2 := "Expected/Value_All".Expected_493)
      Move(in := 493, out1 => #Output)
   END_RUNG
   RUNG wire#powerrail
      { S7_Templates := "SrcType := String" } EQ_Contact(in1 := "Expected/Value_All".V, in2 := "Expected/Value_All".Expected_494)
      Move(in := 494, out1 => #Output)
   END_RUNG
   RUNG wire#powerrail
      { S7_Templates := "SrcType := String" } EQ_Contact(in1 := "Expected/Value_All".V, in2 := "Expected/Value_All".Expected_495)
      Move(in := 495, out1 => #Output)
   END_RUNG
   RUNG wire#powerrail
      { S7_Templates := "SrcType := String" } EQ_Contact(in1 := "Expected/Value_All".V, in2 := "Expected/Value_All".Expected_496)
      Move(in := 496, out1 => #Output)
   END_RUNG
   RUNG wire#powerrail
      { S7_Templates := "SrcType := String" } EQ_Contact(in1 := "Expected/Value_All".V, in2 := "Expected/Value_All".Expected_497)
      Move(in := 497, out1 => #Output)
   END_RUNG
   RUNG wire#powerrail
      { S7_Templates := "SrcType := String" } EQ_Contact(in1 := "Expected/Value_All".V, in2 := "Expected/Value_All".Expected_498)
      Move(in := 498, out1 => #Output)
   END_RUNG
   RUNG wire#powerrail
      { S7_Templates := "SrcType := String" } EQ_Contact(in1 := "Expected/Value_All".V, in2 := "Expected/Value_All".Expected_499)
      Move(in := 499, out1 => #Output)
   END_RUNG
   RUNG wire#powerrail
      { S7_Templates := "SrcType := String" } EQ_Contact(in1 := "Expected/Value_All".V, in2 := "Expected/Value_All".Expected_500)
      Move(in := 500, out1 => #Output)
   END_RUNG
   // the same network as SCL:
   IF "Expected/Value_All".V = "Expected/Value_All".Expected_481 THEN #Output := 481; END_IF;
   IF "Expected/Value_All".V = "Expected/Value_All".Expected_482 THEN #Output := 482; END_IF;
   IF "Expected/Value_All".V = "Expected/Value_All".Expected_483 THEN #Output := 483; END_IF;
   IF "Expected/Value_All".V = "Expected/Value_All".Expected_484 THEN #Output := 484; END_IF;
   IF "Expected/Value_All".V = "Expected/Value_All".Expected_485 THEN #Output := 485; END_IF;
   IF "Expected/Value_All".V = "Expected/Value_All".Expected_486 THEN #Output := 486; END_IF;
   IF "Expected/Value_All".V = "Expected/Value_All".Expected_487 THEN #Output := 487; END_IF;
   IF "Expected/Value_All".V = "Expected/Value_All".Expected_488 THEN #Output := 488; END_IF;
   IF "Expected/Value_All".V = "Expected/Value_All".Expected_489 THEN #Output := 489; END_IF;
   IF "Expected/Value_All".V = "Expected/Value_All".Expected_490 THEN #Output := 490; END_IF;
   IF "Expected/Value_All".V = "Expected/Value_All".Expected_491 THEN #Output := 491; END_IF;
   IF "Expected/Value_All".V = "Expected/Value_All".Expected_492 THEN #Output := 492; END_IF;
   IF "Expected/Value_All".V = "Expected/Value_All".Expected_493 THEN #Output := 493; END_IF;
   IF "Expected/Value_All".V = "Expected/Value_All".Expected_494 THEN #Output := 494; END_IF;
   IF "Expected/Value_All".V = "Expected/Value_All".Expected_495 THEN #Output := 495; END_IF;
   IF "Expected/Value_All".V = "Expected/Value_All".Expected_496 THEN #Output := 496; END_IF;
   IF "Expected/Value_All".V = "Expected/Value_All".Expected_497 THEN #Output := 497; END_IF;
   IF "Expected/Value_All".V = "Expected/Value_All".Expected_498 THEN #Output := 498; END_IF;
   IF "Expected/Value_All".V = "Expected/Value_All".Expected_499 THEN #Output := 499; END_IF;
   IF "Expected/Value_All".V = "Expected/Value_All".Expected_500 THEN #Output := 500; END_IF;
END_REGION

REGION Network 26
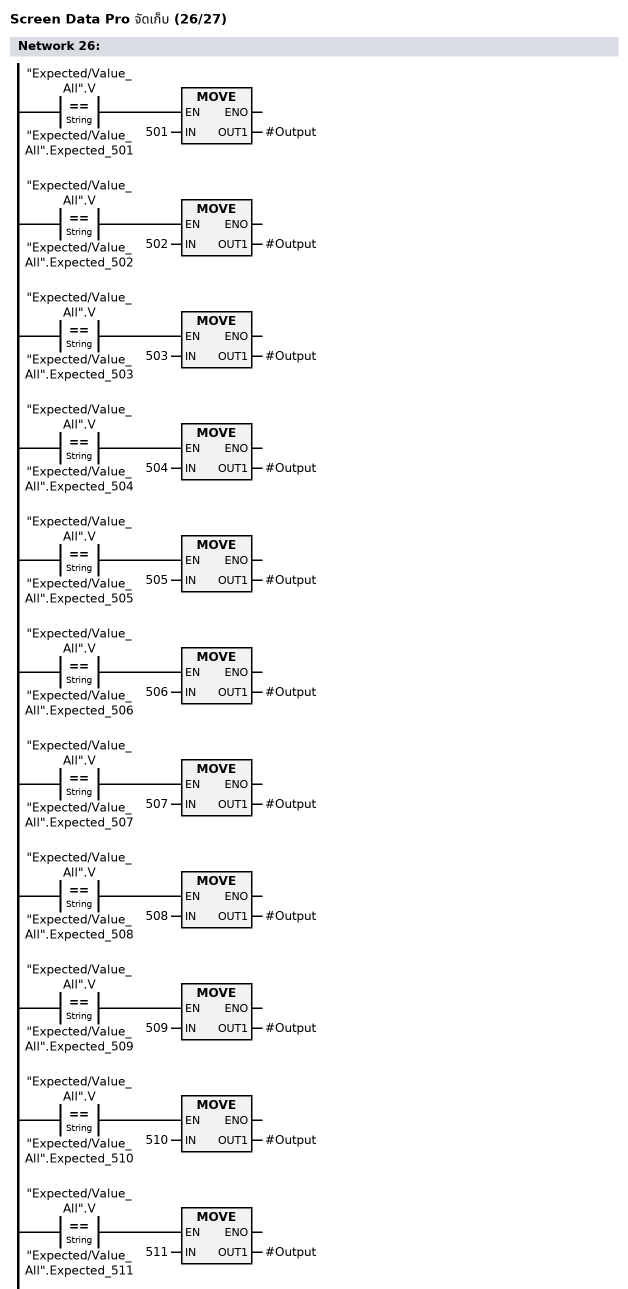
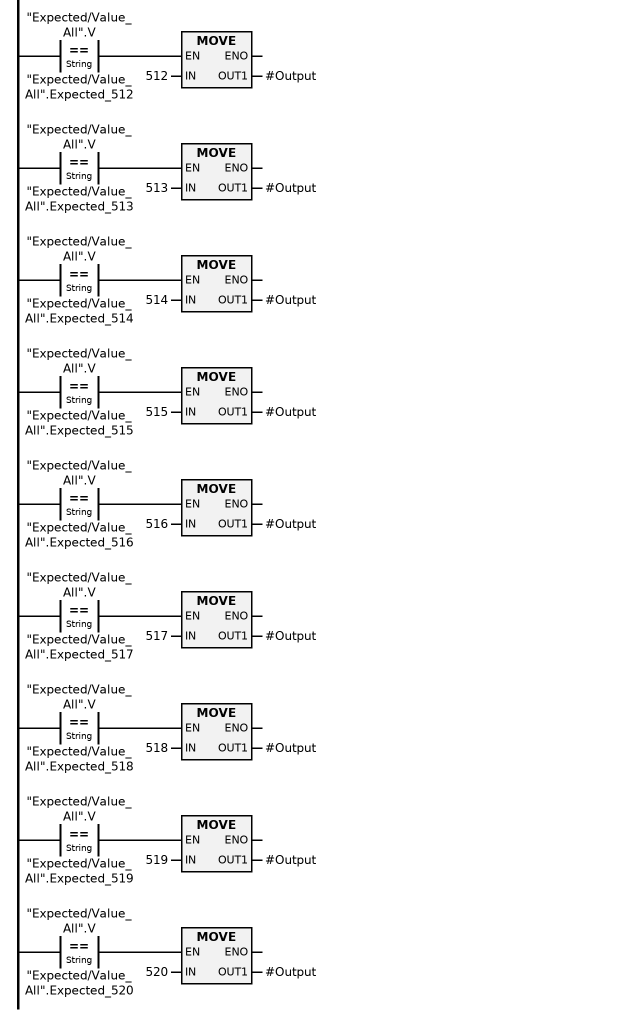
   RUNG wire#powerrail
      { S7_Templates := "SrcType := String" } EQ_Contact(in1 := "Expected/Value_All".V, in2 := "Expected/Value_All".Expected_501)
      Move(in := 501, out1 => #Output)
   END_RUNG
   RUNG wire#powerrail
      { S7_Templates := "SrcType := String" } EQ_Contact(in1 := "Expected/Value_All".V, in2 := "Expected/Value_All".Expected_502)
      Move(in := 502, out1 => #Output)
   END_RUNG
   RUNG wire#powerrail
      { S7_Templates := "SrcType := String" } EQ_Contact(in1 := "Expected/Value_All".V, in2 := "Expected/Value_All".Expected_503)
      Move(in := 503, out1 => #Output)
   END_RUNG
   RUNG wire#powerrail
      { S7_Templates := "SrcType := String" } EQ_Contact(in1 := "Expected/Value_All".V, in2 := "Expected/Value_All".Expected_504)
      Move(in := 504, out1 => #Output)
   END_RUNG
   RUNG wire#powerrail
      { S7_Templates := "SrcType := String" } EQ_Contact(in1 := "Expected/Value_All".V, in2 := "Expected/Value_All".Expected_505)
      Move(in := 505, out1 => #Output)
   END_RUNG
   RUNG wire#powerrail
      { S7_Templates := "SrcType := String" } EQ_Contact(in1 := "Expected/Value_All".V, in2 := "Expected/Value_All".Expected_506)
      Move(in := 506, out1 => #Output)
   END_RUNG
   RUNG wire#powerrail
      { S7_Templates := "SrcType := String" } EQ_Contact(in1 := "Expected/Value_All".V, in2 := "Expected/Value_All".Expected_507)
      Move(in := 507, out1 => #Output)
   END_RUNG
   RUNG wire#powerrail
      { S7_Templates := "SrcType := String" } EQ_Contact(in1 := "Expected/Value_All".V, in2 := "Expected/Value_All".Expected_508)
      Move(in := 508, out1 => #Output)
   END_RUNG
   RUNG wire#powerrail
      { S7_Templates := "SrcType := String" } EQ_Contact(in1 := "Expected/Value_All".V, in2 := "Expected/Value_All".Expected_509)
      Move(in := 509, out1 => #Output)
   END_RUNG
   RUNG wire#powerrail
      { S7_Templates := "SrcType := String" } EQ_Contact(in1 := "Expected/Value_All".V, in2 := "Expected/Value_All".Expected_510)
      Move(in := 510, out1 => #Output)
   END_RUNG
   RUNG wire#powerrail
      { S7_Templates := "SrcType := String" } EQ_Contact(in1 := "Expected/Value_All".V, in2 := "Expected/Value_All".Expected_511)
      Move(in := 511, out1 => #Output)
   END_RUNG
   RUNG wire#powerrail
      { S7_Templates := "SrcType := String" } EQ_Contact(in1 := "Expected/Value_All".V, in2 := "Expected/Value_All".Expected_512)
      Move(in := 512, out1 => #Output)
   END_RUNG
   RUNG wire#powerrail
      { S7_Templates := "SrcType := String" } EQ_Contact(in1 := "Expected/Value_All".V, in2 := "Expected/Value_All".Expected_513)
      Move(in := 513, out1 => #Output)
   END_RUNG
   RUNG wire#powerrail
      { S7_Templates := "SrcType := String" } EQ_Contact(in1 := "Expected/Value_All".V, in2 := "Expected/Value_All".Expected_514)
      Move(in := 514, out1 => #Output)
   END_RUNG
   RUNG wire#powerrail
      { S7_Templates := "SrcType := String" } EQ_Contact(in1 := "Expected/Value_All".V, in2 := "Expected/Value_All".Expected_515)
      Move(in := 515, out1 => #Output)
   END_RUNG
   RUNG wire#powerrail
      { S7_Templates := "SrcType := String" } EQ_Contact(in1 := "Expected/Value_All".V, in2 := "Expected/Value_All".Expected_516)
      Move(in := 516, out1 => #Output)
   END_RUNG
   RUNG wire#powerrail
      { S7_Templates := "SrcType := String" } EQ_Contact(in1 := "Expected/Value_All".V, in2 := "Expected/Value_All".Expected_517)
      Move(in := 517, out1 => #Output)
   END_RUNG
   RUNG wire#powerrail
      { S7_Templates := "SrcType := String" } EQ_Contact(in1 := "Expected/Value_All".V, in2 := "Expected/Value_All".Expected_518)
      Move(in := 518, out1 => #Output)
   END_RUNG
   RUNG wire#powerrail
      { S7_Templates := "SrcType := String" } EQ_Contact(in1 := "Expected/Value_All".V, in2 := "Expected/Value_All".Expected_519)
      Move(in := 519, out1 => #Output)
   END_RUNG
   RUNG wire#powerrail
      { S7_Templates := "SrcType := String" } EQ_Contact(in1 := "Expected/Value_All".V, in2 := "Expected/Value_All".Expected_520)
      Move(in := 520, out1 => #Output)
   END_RUNG
   // the same network as SCL:
   IF "Expected/Value_All".V = "Expected/Value_All".Expected_501 THEN #Output := 501; END_IF;
   IF "Expected/Value_All".V = "Expected/Value_All".Expected_502 THEN #Output := 502; END_IF;
   IF "Expected/Value_All".V = "Expected/Value_All".Expected_503 THEN #Output := 503; END_IF;
   IF "Expected/Value_All".V = "Expected/Value_All".Expected_504 THEN #Output := 504; END_IF;
   IF "Expected/Value_All".V = "Expected/Value_All".Expected_505 THEN #Output := 505; END_IF;
   IF "Expected/Value_All".V = "Expected/Value_All".Expected_506 THEN #Output := 506; END_IF;
   IF "Expected/Value_All".V = "Expected/Value_All".Expected_507 THEN #Output := 507; END_IF;
   IF "Expected/Value_All".V = "Expected/Value_All".Expected_508 THEN #Output := 508; END_IF;
   IF "Expected/Value_All".V = "Expected/Value_All".Expected_509 THEN #Output := 509; END_IF;
   IF "Expected/Value_All".V = "Expected/Value_All".Expected_510 THEN #Output := 510; END_IF;
   IF "Expected/Value_All".V = "Expected/Value_All".Expected_511 THEN #Output := 511; END_IF;
   IF "Expected/Value_All".V = "Expected/Value_All".Expected_512 THEN #Output := 512; END_IF;
   IF "Expected/Value_All".V = "Expected/Value_All".Expected_513 THEN #Output := 513; END_IF;
   IF "Expected/Value_All".V = "Expected/Value_All".Expected_514 THEN #Output := 514; END_IF;
   IF "Expected/Value_All".V = "Expected/Value_All".Expected_515 THEN #Output := 515; END_IF;
   IF "Expected/Value_All".V = "Expected/Value_All".Expected_516 THEN #Output := 516; END_IF;
   IF "Expected/Value_All".V = "Expected/Value_All".Expected_517 THEN #Output := 517; END_IF;
   IF "Expected/Value_All".V = "Expected/Value_All".Expected_518 THEN #Output := 518; END_IF;
   IF "Expected/Value_All".V = "Expected/Value_All".Expected_519 THEN #Output := 519; END_IF;
   IF "Expected/Value_All".V = "Expected/Value_All".Expected_520 THEN #Output := 520; END_IF;
END_REGION

REGION Network 27
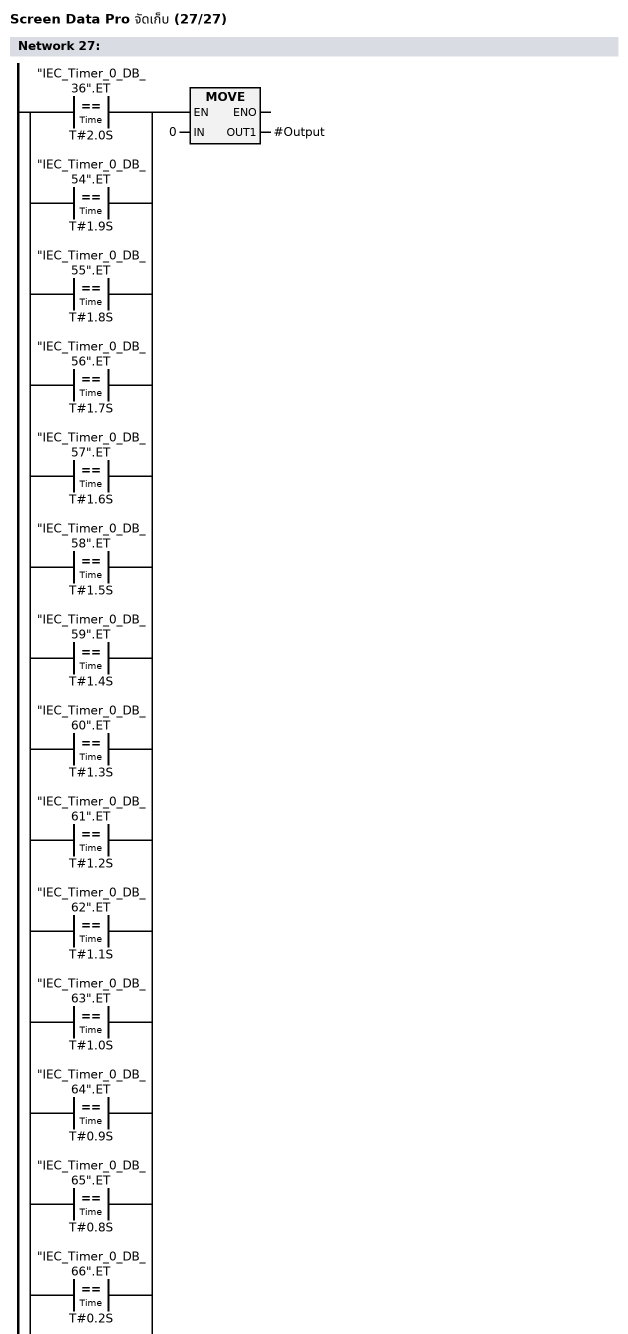
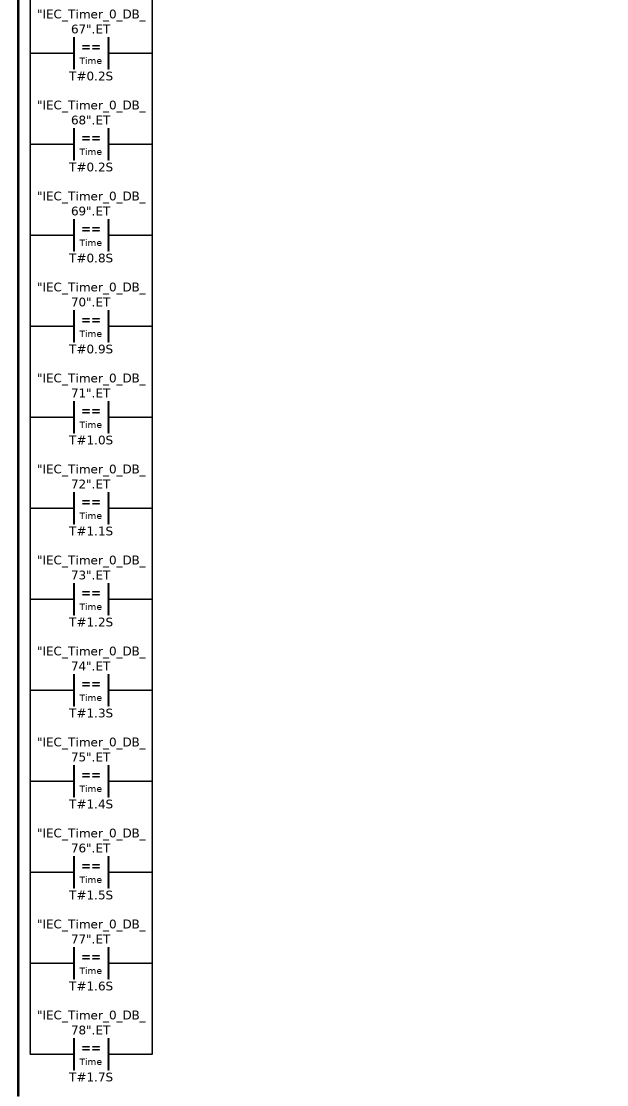
   RUNG wire#powerrail
      { S7_Templates := "SrcType := Time" } EQ_Contact(in1 := "IEC_Timer_0_DB_36".ET, in2 := T#2.0S)
      wire#w1
      Move(in := 0, out1 => #Output)
   END_RUNG
   RUNG wire#powerrail
      { S7_Templates := "SrcType := Time" } EQ_Contact(in1 := "IEC_Timer_0_DB_54".ET, in2 := T#1.9S)
   END_RUNG wire#w1
   RUNG wire#powerrail
      { S7_Templates := "SrcType := Time" } EQ_Contact(in1 := "IEC_Timer_0_DB_55".ET, in2 := T#1.8S)
   END_RUNG wire#w1
   RUNG wire#powerrail
      { S7_Templates := "SrcType := Time" } EQ_Contact(in1 := "IEC_Timer_0_DB_56".ET, in2 := T#1.7S)
   END_RUNG wire#w1
   RUNG wire#powerrail
      { S7_Templates := "SrcType := Time" } EQ_Contact(in1 := "IEC_Timer_0_DB_57".ET, in2 := T#1.6S)
   END_RUNG wire#w1
   RUNG wire#powerrail
      { S7_Templates := "SrcType := Time" } EQ_Contact(in1 := "IEC_Timer_0_DB_58".ET, in2 := T#1.5S)
   END_RUNG wire#w1
   RUNG wire#powerrail
      { S7_Templates := "SrcType := Time" } EQ_Contact(in1 := "IEC_Timer_0_DB_59".ET, in2 := T#1.4S)
   END_RUNG wire#w1
   RUNG wire#powerrail
      { S7_Templates := "SrcType := Time" } EQ_Contact(in1 := "IEC_Timer_0_DB_60".ET, in2 := T#1.3S)
   END_RUNG wire#w1
   RUNG wire#powerrail
      { S7_Templates := "SrcType := Time" } EQ_Contact(in1 := "IEC_Timer_0_DB_61".ET, in2 := T#1.2S)
   END_RUNG wire#w1
   RUNG wire#powerrail
      { S7_Templates := "SrcType := Time" } EQ_Contact(in1 := "IEC_Timer_0_DB_62".ET, in2 := T#1.1S)
   END_RUNG wire#w1
   RUNG wire#powerrail
      { S7_Templates := "SrcType := Time" } EQ_Contact(in1 := "IEC_Timer_0_DB_63".ET, in2 := T#1.0S)
   END_RUNG wire#w1
   RUNG wire#powerrail
      { S7_Templates := "SrcType := Time" } EQ_Contact(in1 := "IEC_Timer_0_DB_64".ET, in2 := T#0.9S)
   END_RUNG wire#w1
   RUNG wire#powerrail
      { S7_Templates := "SrcType := Time" } EQ_Contact(in1 := "IEC_Timer_0_DB_65".ET, in2 := T#0.8S)
   END_RUNG wire#w1
   RUNG wire#powerrail
      { S7_Templates := "SrcType := Time" } EQ_Contact(in1 := "IEC_Timer_0_DB_66".ET, in2 := T#0.2S)
   END_RUNG wire#w1
   RUNG wire#powerrail
      { S7_Templates := "SrcType := Time" } EQ_Contact(in1 := "IEC_Timer_0_DB_67".ET, in2 := T#0.2S)
   END_RUNG wire#w1
   RUNG wire#powerrail
      { S7_Templates := "SrcType := Time" } EQ_Contact(in1 := "IEC_Timer_0_DB_68".ET, in2 := T#0.2S)
   END_RUNG wire#w1
   RUNG wire#powerrail
      { S7_Templates := "SrcType := Time" } EQ_Contact(in1 := "IEC_Timer_0_DB_69".ET, in2 := T#0.8S)
   END_RUNG wire#w1
   RUNG wire#powerrail
      { S7_Templates := "SrcType := Time" } EQ_Contact(in1 := "IEC_Timer_0_DB_70".ET, in2 := T#0.9S)
   END_RUNG wire#w1
   RUNG wire#powerrail
      { S7_Templates := "SrcType := Time" } EQ_Contact(in1 := "IEC_Timer_0_DB_71".ET, in2 := T#1.0S)
   END_RUNG wire#w1
   RUNG wire#powerrail
      { S7_Templates := "SrcType := Time" } EQ_Contact(in1 := "IEC_Timer_0_DB_72".ET, in2 := T#1.1S)
   END_RUNG wire#w1
   RUNG wire#powerrail
      { S7_Templates := "SrcType := Time" } EQ_Contact(in1 := "IEC_Timer_0_DB_73".ET, in2 := T#1.2S)
   END_RUNG wire#w1
   RUNG wire#powerrail
      { S7_Templates := "SrcType := Time" } EQ_Contact(in1 := "IEC_Timer_0_DB_74".ET, in2 := T#1.3S)
   END_RUNG wire#w1
   RUNG wire#powerrail
      { S7_Templates := "SrcType := Time" } EQ_Contact(in1 := "IEC_Timer_0_DB_75".ET, in2 := T#1.4S)
   END_RUNG wire#w1
   RUNG wire#powerrail
      { S7_Templates := "SrcType := Time" } EQ_Contact(in1 := "IEC_Timer_0_DB_76".ET, in2 := T#1.5S)
   END_RUNG wire#w1
   RUNG wire#powerrail
      { S7_Templates := "SrcType := Time" } EQ_Contact(in1 := "IEC_Timer_0_DB_77".ET, in2 := T#1.6S)
   END_RUNG wire#w1
   RUNG wire#powerrail
      { S7_Templates := "SrcType := Time" } EQ_Contact(in1 := "IEC_Timer_0_DB_78".ET, in2 := T#1.7S)
   END_RUNG wire#w1
   // the same network as SCL:
   IF ("IEC_Timer_0_DB_36".ET = T#2.0S) OR ("IEC_Timer_0_DB_54".ET = T#1.9S) OR ("IEC_Timer_0_DB_55".ET = T#1.8S) OR ("IEC_Timer_0_DB_56".ET = T#1.7S) OR ("IEC_Timer_0_DB_57".ET = T#1.6S) OR ("IEC_Timer_0_DB_58".ET = T#1.5S) OR ("IEC_Timer_0_DB_59".ET = T#1.4S) OR ("IEC_Timer_0_DB_60".ET = T#1.3S) OR ("IEC_Timer_0_DB_61".ET = T#1.2S) OR ("IEC_Timer_0_DB_62".ET = T#1.1S) OR ("IEC_Timer_0_DB_63".ET = T#1.0S) OR ("IEC_Timer_0_DB_64".ET = T#0.9S) OR ("IEC_Timer_0_DB_65".ET = T#0.8S) OR ("IEC_Timer_0_DB_66".ET = T#0.2S) OR ("IEC_Timer_0_DB_67".ET = T#0.2S) OR ("IEC_Timer_0_DB_68".ET = T#0.2S) OR ("IEC_Timer_0_DB_69".ET = T#0.8S) OR ("IEC_Timer_0_DB_70".ET = T#0.9S) OR ("IEC_Timer_0_DB_71".ET = T#1.0S) OR ("IEC_Timer_0_DB_72".ET = T#1.1S) OR ("IEC_Timer_0_DB_73".ET = T#1.2S) OR ("IEC_Timer_0_DB_74".ET = T#1.3S) OR ("IEC_Timer_0_DB_75".ET = T#1.4S) OR ("IEC_Timer_0_DB_76".ET = T#1.5S) OR ("IEC_Timer_0_DB_77".ET = T#1.6S) OR ("IEC_Timer_0_DB_78".ET = T#1.7S) THEN
       #Output := 0;
   END_IF;
END_REGION
END_FUNCTION_BLOCK

FUNCTION_BLOCK "บันทึกผลการเคลื่อนที่ ไว้ที่ Excell"   // FB12, LAD
{ S7_Optimized_Access := 'TRUE' }
VERSION : 0.1
   VAR
      Alarms : Word;
   END_VAR
BEGIN

REGION Network 1: Alarms
   // Motor
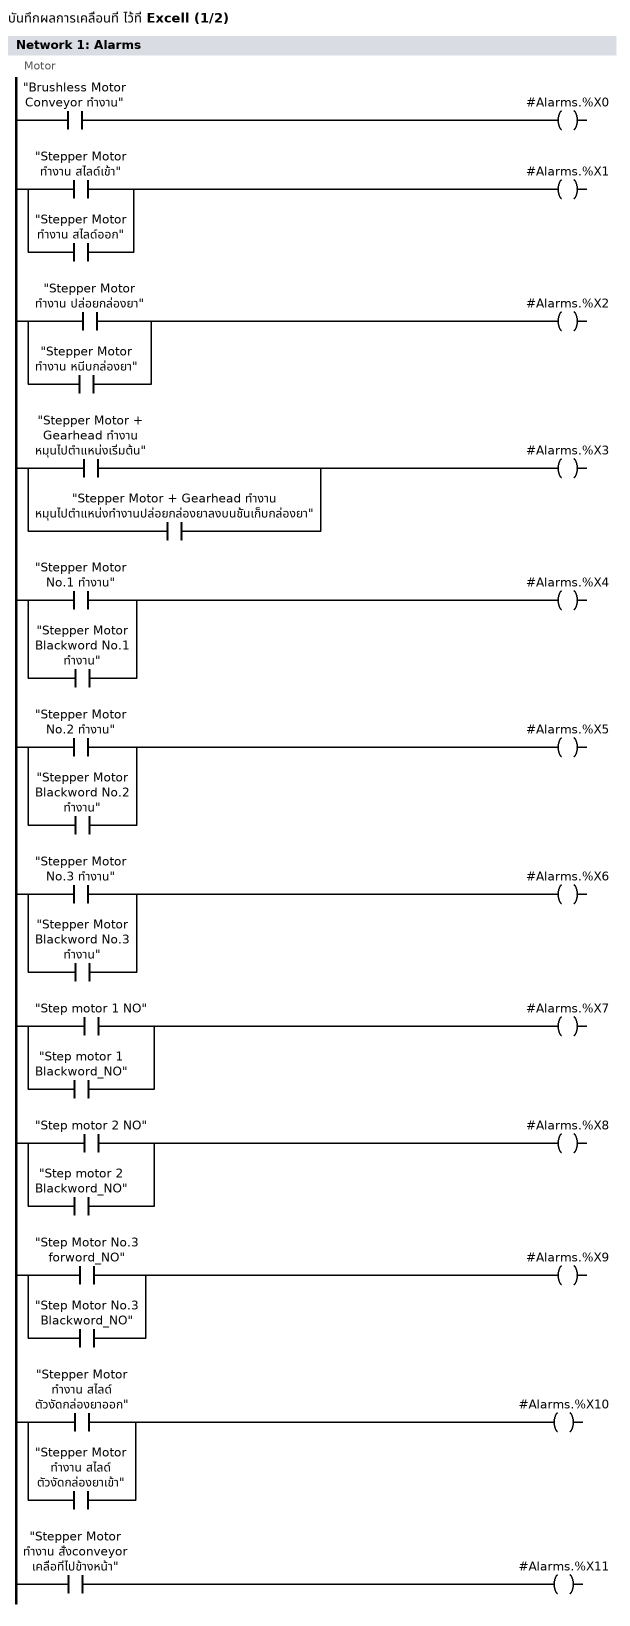
   RUNG wire#powerrail
      Contact( "Brushless Motor Conveyor ทำงาน" )
      Coil( #Alarms.%X0 )
   END_RUNG
   RUNG wire#powerrail
      Contact( "Stepper Motor ทำงาน สไลด์เข้า" )
      wire#w1
      Coil( #Alarms.%X1 )
   END_RUNG
   RUNG wire#powerrail
      Contact( "Stepper Motor ทำงาน สไลด์ออก" )
   END_RUNG wire#w1
   RUNG wire#powerrail
      Contact( "Stepper Motor ทำงาน ปล่อยกล่องยา" )
      wire#w2
      Coil( #Alarms.%X2 )
   END_RUNG
   RUNG wire#powerrail
      Contact( "Stepper Motor ทำงาน หนีบกล่องยา" )
   END_RUNG wire#w2
   RUNG wire#powerrail
      Contact( "Stepper Motor + Gearhead ทำงาน หมุนไปตำแหน่งเริ่มต้น" )
      wire#w3
      Coil( #Alarms.%X3 )
   END_RUNG
   RUNG wire#powerrail
      Contact( "Stepper Motor + Gearhead ทำงาน หมุนไปตำแหน่งทำงานปล่อยกล่องยาลงบนชั้นเก็บกล่องยา" )
   END_RUNG wire#w3
   RUNG wire#powerrail
      Contact( "Stepper Motor No.1 ทำงาน" )
      wire#w4
      Coil( #Alarms.%X4 )
   END_RUNG
   RUNG wire#powerrail
      Contact( "Stepper Motor Blackword No.1 ทำงาน" )
   END_RUNG wire#w4
   RUNG wire#powerrail
      Contact( "Stepper Motor No.2 ทำงาน" )
      wire#w5
      Coil( #Alarms.%X5 )
   END_RUNG
   RUNG wire#powerrail
      Contact( "Stepper Motor Blackword No.2 ทำงาน" )
   END_RUNG wire#w5
   RUNG wire#powerrail
      Contact( "Stepper Motor No.3 ทำงาน" )
      wire#w6
      Coil( #Alarms.%X6 )
   END_RUNG
   RUNG wire#powerrail
      Contact( "Stepper Motor Blackword No.3 ทำงาน" )
   END_RUNG wire#w6
   RUNG wire#powerrail
      Contact( "Step motor 1 NO" )
      wire#w7
      Coil( #Alarms.%X7 )
   END_RUNG
   RUNG wire#powerrail
      Contact( "Step motor 1 Blackword_NO" )
   END_RUNG wire#w7
   RUNG wire#powerrail
      Contact( "Step motor 2 NO" )
      wire#w8
      Coil( #Alarms.%X8 )
   END_RUNG
   RUNG wire#powerrail
      Contact( "Step motor 2 Blackword_NO" )
   END_RUNG wire#w8
   RUNG wire#powerrail
      Contact( "Step Motor No.3 forword_NO" )
      wire#w9
      Coil( #Alarms.%X9 )
   END_RUNG
   RUNG wire#powerrail
      Contact( "Step Motor No.3 Blackword_NO" )
   END_RUNG wire#w9
   RUNG wire#powerrail
      Contact( "Stepper Motor ทำงาน สไลด์ ตัวงัดกล่องยาออก" )
      wire#w10
      Coil( #Alarms.%X10 )
   END_RUNG
   RUNG wire#powerrail
      Contact( "Stepper Motor ทำงาน สไลด์ ตัวงัดกล่องยาเข้า" )
   END_RUNG wire#w10
   RUNG wire#powerrail
      Contact( "Stepper Motor ทำงาน สั่งconveyor เคลื่อที่ไปข้างหน้า" )
      Coil( #Alarms.%X11 )
   END_RUNG
   // the same network as SCL:
   #Alarms.%X0 := "Brushless Motor Conveyor ทำงาน";
   #Alarms.%X1 := "Stepper Motor ทำงาน สไลด์เข้า" OR "Stepper Motor ทำงาน สไลด์ออก";
   #Alarms.%X2 := "Stepper Motor ทำงาน ปล่อยกล่องยา" OR "Stepper Motor ทำงาน หนีบกล่องยา";
   #Alarms.%X3 := "Stepper Motor + Gearhead ทำงาน หมุนไปตำแหน่งเริ่มต้น" OR "Stepper Motor + Gearhead ทำงาน หมุนไปตำแหน่งทำงานปล่อยกล่องยาลงบนชั้นเก็บกล่องยา";
   #Alarms.%X4 := "Stepper Motor No.1 ทำงาน" OR "Stepper Motor Blackword No.1 ทำงาน";
   #Alarms.%X5 := "Stepper Motor No.2 ทำงาน" OR "Stepper Motor Blackword No.2 ทำงาน";
   #Alarms.%X6 := "Stepper Motor No.3 ทำงาน" OR "Stepper Motor Blackword No.3 ทำงาน";
   #Alarms.%X7 := "Step motor 1 NO" OR "Step motor 1 Blackword_NO";
   #Alarms.%X8 := "Step motor 2 NO" OR "Step motor 2 Blackword_NO";
   #Alarms.%X9 := "Step Motor No.3 forword_NO" OR "Step Motor No.3 Blackword_NO";
   #Alarms.%X10 := "Stepper Motor ทำงาน สไลด์ ตัวงัดกล่องยาออก" OR "Stepper Motor ทำงาน สไลด์ ตัวงัดกล่องยาเข้า";
   #Alarms.%X11 := "Stepper Motor ทำงาน สั่งconveyor เคลื่อที่ไปข้างหน้า";
END_REGION

REGION Network 2
   // Sensor (จัดเก็บ)
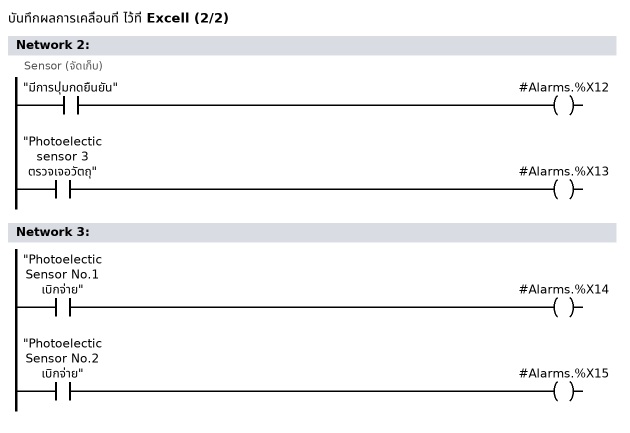
   RUNG wire#powerrail
      Contact( "มีการปุ่มกดยืนยัน" )
      Coil( #Alarms.%X12 )
   END_RUNG
   RUNG wire#powerrail
      Contact( "Photoelectic sensor 3 ตรวจเจอวัตถุ" )
      Coil( #Alarms.%X13 )
   END_RUNG
   // the same network as SCL:
   #Alarms.%X12 := "มีการปุ่มกดยืนยัน";
   #Alarms.%X13 := "Photoelectic sensor 3 ตรวจเจอวัตถุ";
END_REGION

REGION Network 3
   RUNG wire#powerrail
      Contact( "Photoelectic Sensor No.1 เบิกจ่าย" )
      Coil( #Alarms.%X14 )
   END_RUNG
   RUNG wire#powerrail
      Contact( "Photoelectic Sensor No.2 เบิกจ่าย" )
      Coil( #Alarms.%X15 )
   END_RUNG
   // the same network as SCL:
   #Alarms.%X14 := "Photoelectic Sensor No.1 เบิกจ่าย";
   #Alarms.%X15 := "Photoelectic Sensor No.2 เบิกจ่าย";
END_REGION
END_FUNCTION_BLOCK

FUNCTION "Screen 1" : Void   // FC13, LAD
{ S7_Optimized_Access := 'TRUE' }
VERSION : 0.1
BEGIN

REGION Network 1
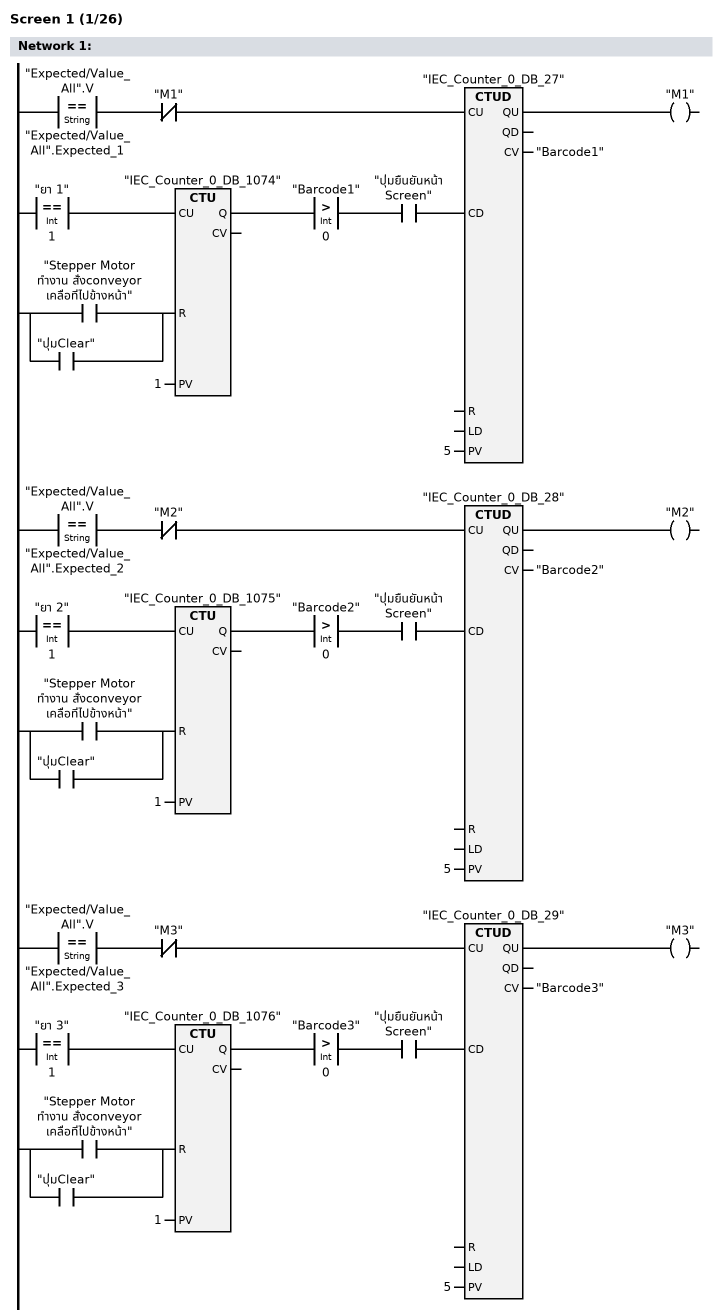
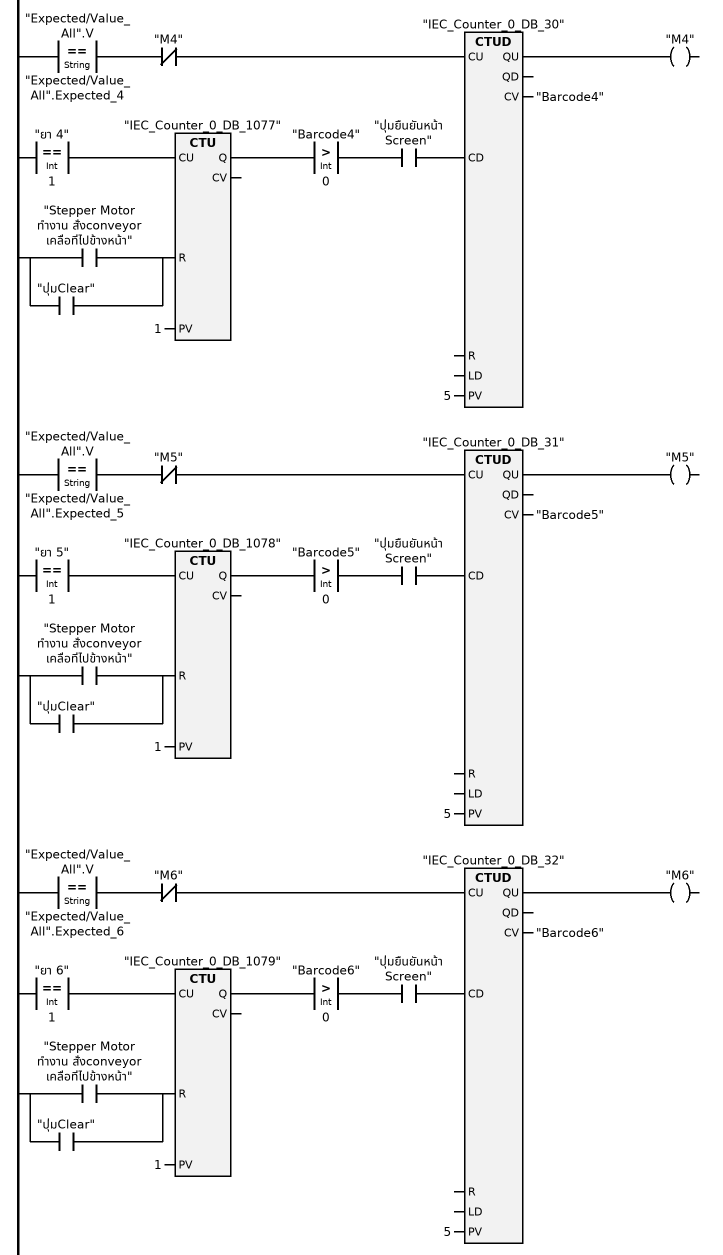
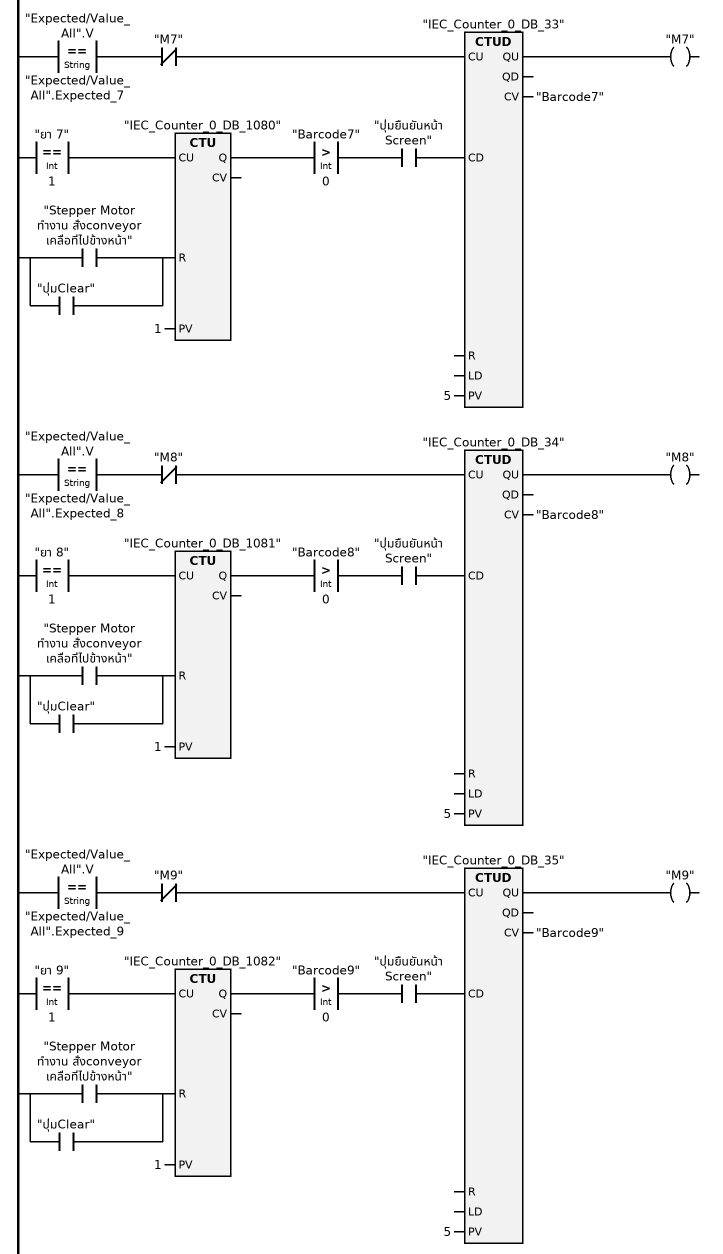
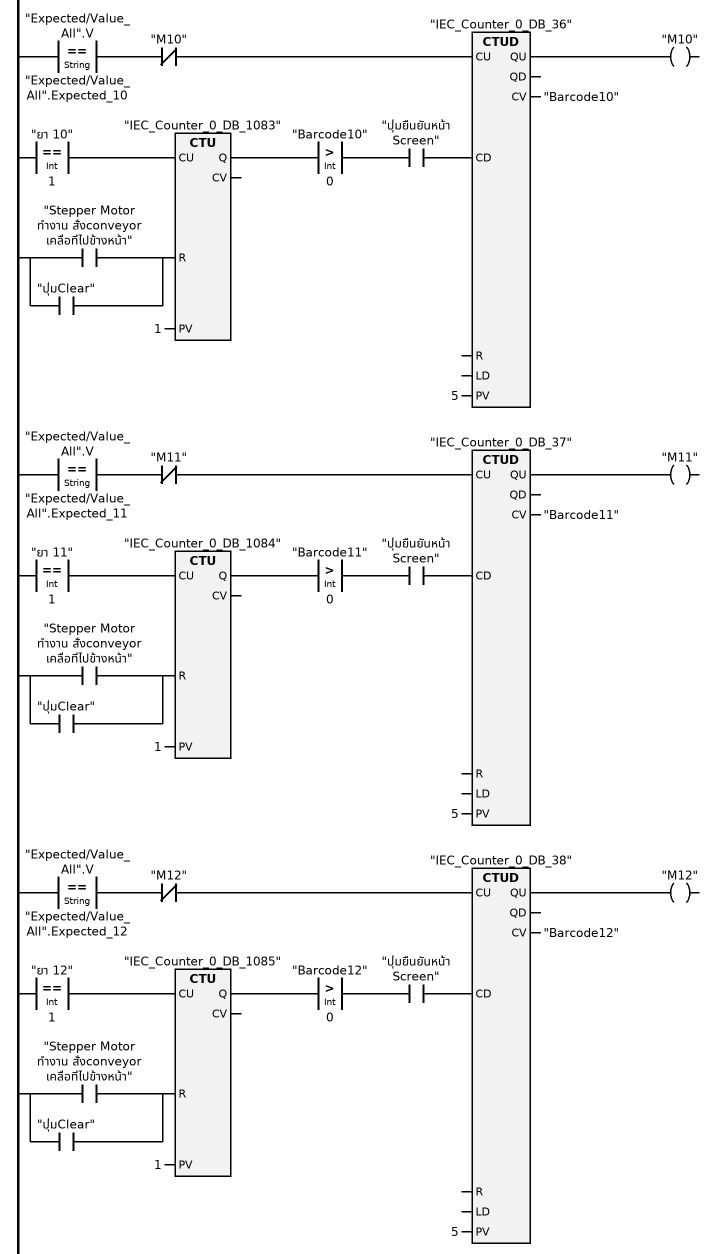
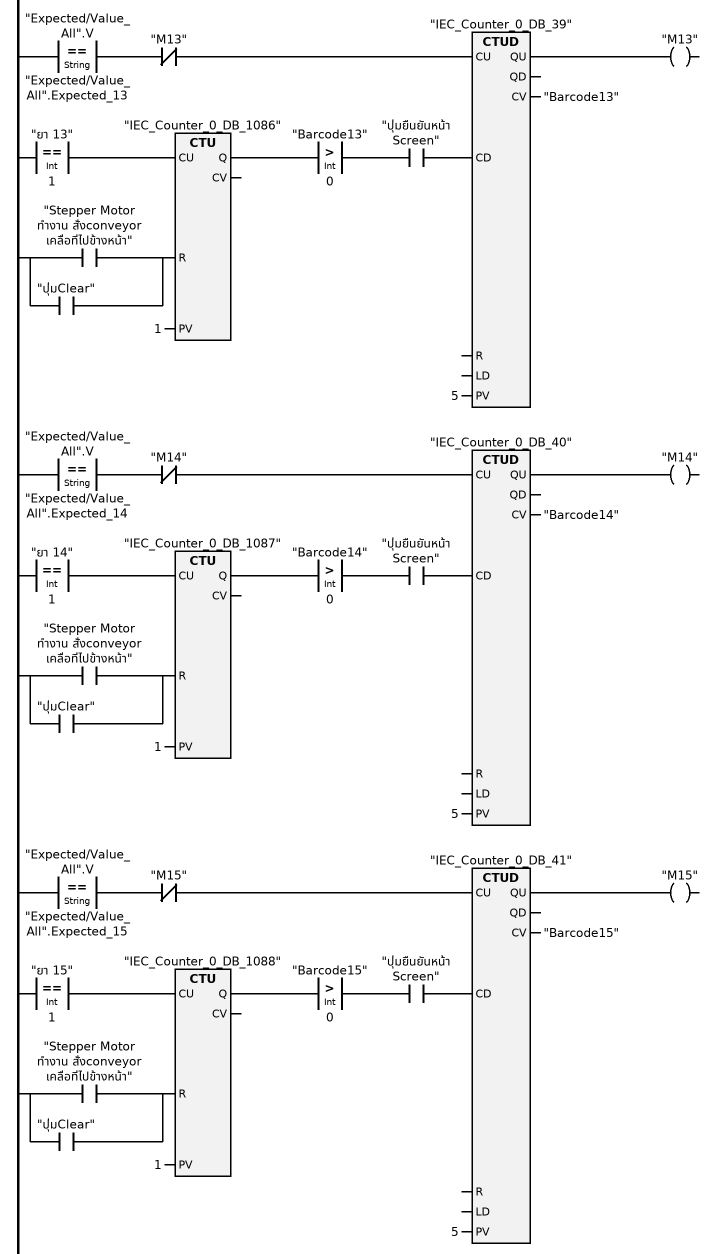
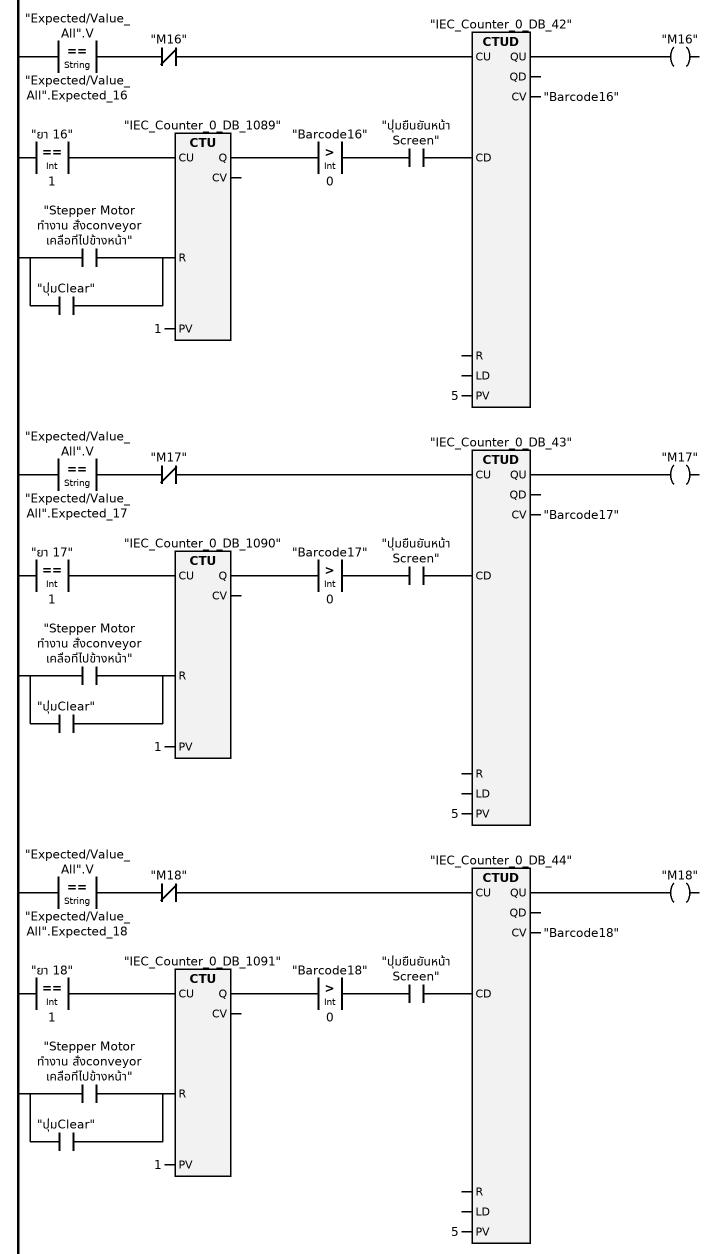
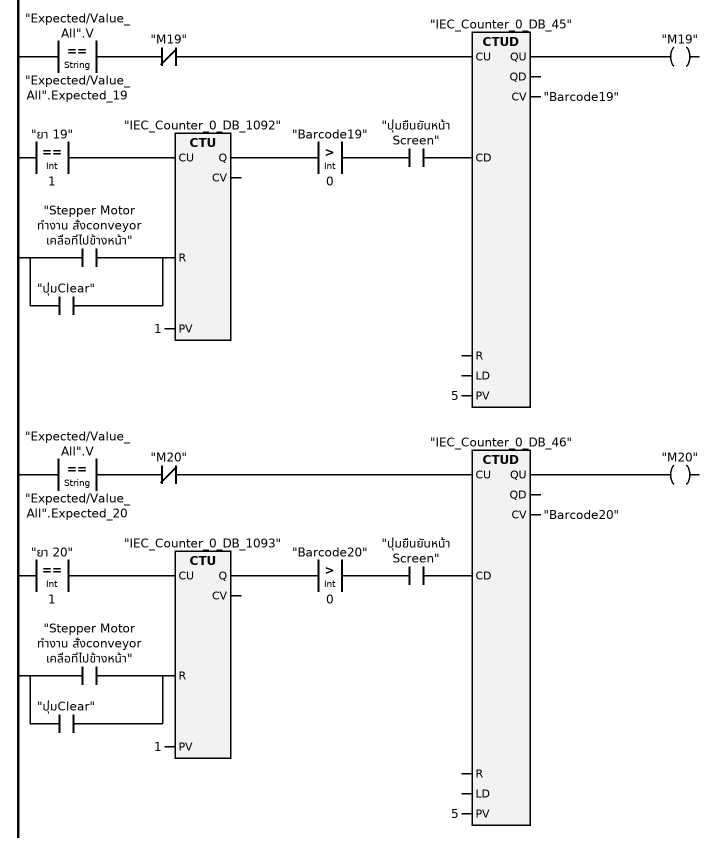
   "IEC_Counter_0_DB_1074".CTU(CU := "ยา 1" = 1,
                           R := "Stepper Motor ทำงาน สั่งconveyor เคลื่อที่ไปข้างหน้า" OR "ปุ่มClear",
                           PV := 1);
   "IEC_Counter_0_DB_27".CTUD(CU := ("Expected/Value_All".V = "Expected/Value_All".Expected_1) AND NOT "M1",
                           CD := "IEC_Counter_0_DB_1074".Q AND ("Barcode1" > 0) AND "ปุ่มยืนยันหน้า Screen",
                           PV := 5,
                           CV => "Barcode1");
   "M1" := "IEC_Counter_0_DB_27".QU;
   "IEC_Counter_0_DB_1075".CTU(CU := "ยา 2" = 1,
                           R := "Stepper Motor ทำงาน สั่งconveyor เคลื่อที่ไปข้างหน้า" OR "ปุ่มClear",
                           PV := 1);
   "IEC_Counter_0_DB_28".CTUD(CU := ("Expected/Value_All".V = "Expected/Value_All".Expected_2) AND NOT "M2",
                           CD := "IEC_Counter_0_DB_1075".Q AND ("Barcode2" > 0) AND "ปุ่มยืนยันหน้า Screen",
                           PV := 5,
                           CV => "Barcode2");
   "M2" := "IEC_Counter_0_DB_28".QU;
   "IEC_Counter_0_DB_1076".CTU(CU := "ยา 3" = 1,
                           R := "Stepper Motor ทำงาน สั่งconveyor เคลื่อที่ไปข้างหน้า" OR "ปุ่มClear",
                           PV := 1);
   "IEC_Counter_0_DB_29".CTUD(CU := ("Expected/Value_All".V = "Expected/Value_All".Expected_3) AND NOT "M3",
                           CD := "IEC_Counter_0_DB_1076".Q AND ("Barcode3" > 0) AND "ปุ่มยืนยันหน้า Screen",
                           PV := 5,
                           CV => "Barcode3");
   "M3" := "IEC_Counter_0_DB_29".QU;
   "IEC_Counter_0_DB_1077".CTU(CU := "ยา 4" = 1,
                           R := "Stepper Motor ทำงาน สั่งconveyor เคลื่อที่ไปข้างหน้า" OR "ปุ่มClear",
                           PV := 1);
   "IEC_Counter_0_DB_30".CTUD(CU := ("Expected/Value_All".V = "Expected/Value_All".Expected_4) AND NOT "M4",
                           CD := "IEC_Counter_0_DB_1077".Q AND ("Barcode4" > 0) AND "ปุ่มยืนยันหน้า Screen",
                           PV := 5,
                           CV => "Barcode4");
   "M4" := "IEC_Counter_0_DB_30".QU;
   "IEC_Counter_0_DB_1078".CTU(CU := "ยา 5" = 1,
                           R := "Stepper Motor ทำงาน สั่งconveyor เคลื่อที่ไปข้างหน้า" OR "ปุ่มClear",
                           PV := 1);
   "IEC_Counter_0_DB_31".CTUD(CU := ("Expected/Value_All".V = "Expected/Value_All".Expected_5) AND NOT "M5",
                           CD := "IEC_Counter_0_DB_1078".Q AND ("Barcode5" > 0) AND "ปุ่มยืนยันหน้า Screen",
                           PV := 5,
                           CV => "Barcode5");
   "M5" := "IEC_Counter_0_DB_31".QU;
   "IEC_Counter_0_DB_1079".CTU(CU := "ยา 6" = 1,
                           R := "Stepper Motor ทำงาน สั่งconveyor เคลื่อที่ไปข้างหน้า" OR "ปุ่มClear",
                           PV := 1);
   "IEC_Counter_0_DB_32".CTUD(CU := ("Expected/Value_All".V = "Expected/Value_All".Expected_6) AND NOT "M6",
                           CD := "IEC_Counter_0_DB_1079".Q AND ("Barcode6" > 0) AND "ปุ่มยืนยันหน้า Screen",
                           PV := 5,
                           CV => "Barcode6");
   "M6" := "IEC_Counter_0_DB_32".QU;
   "IEC_Counter_0_DB_1080".CTU(CU := "ยา 7" = 1,
                           R := "Stepper Motor ทำงาน สั่งconveyor เคลื่อที่ไปข้างหน้า" OR "ปุ่มClear",
                           PV := 1);
   "IEC_Counter_0_DB_33".CTUD(CU := ("Expected/Value_All".V = "Expected/Value_All".Expected_7) AND NOT "M7",
                           CD := "IEC_Counter_0_DB_1080".Q AND ("Barcode7" > 0) AND "ปุ่มยืนยันหน้า Screen",
                           PV := 5,
                           CV => "Barcode7");
   "M7" := "IEC_Counter_0_DB_33".QU;
   "IEC_Counter_0_DB_1081".CTU(CU := "ยา 8" = 1,
                           R := "Stepper Motor ทำงาน สั่งconveyor เคลื่อที่ไปข้างหน้า" OR "ปุ่มClear",
                           PV := 1);
   "IEC_Counter_0_DB_34".CTUD(CU := ("Expected/Value_All".V = "Expected/Value_All".Expected_8) AND NOT "M8",
                           CD := "IEC_Counter_0_DB_1081".Q AND ("Barcode8" > 0) AND "ปุ่มยืนยันหน้า Screen",
                           PV := 5,
                           CV => "Barcode8");
   "M8" := "IEC_Counter_0_DB_34".QU;
   "IEC_Counter_0_DB_1082".CTU(CU := "ยา 9" = 1,
                           R := "Stepper Motor ทำงาน สั่งconveyor เคลื่อที่ไปข้างหน้า" OR "ปุ่มClear",
                           PV := 1);
   "IEC_Counter_0_DB_35".CTUD(CU := ("Expected/Value_All".V = "Expected/Value_All".Expected_9) AND NOT "M9",
                           CD := "IEC_Counter_0_DB_1082".Q AND ("Barcode9" > 0) AND "ปุ่มยืนยันหน้า Screen",
                           PV := 5,
                           CV => "Barcode9");
   "M9" := "IEC_Counter_0_DB_35".QU;
   "IEC_Counter_0_DB_1083".CTU(CU := "ยา 10" = 1,
                           R := "Stepper Motor ทำงาน สั่งconveyor เคลื่อที่ไปข้างหน้า" OR "ปุ่มClear",
                           PV := 1);
   "IEC_Counter_0_DB_36".CTUD(CU := ("Expected/Value_All".V = "Expected/Value_All".Expected_10) AND NOT "M10",
                           CD := "IEC_Counter_0_DB_1083".Q AND ("Barcode10" > 0) AND "ปุ่มยืนยันหน้า Screen",
                           PV := 5,
                           CV => "Barcode10");
   "M10" := "IEC_Counter_0_DB_36".QU;
   "IEC_Counter_0_DB_1084".CTU(CU := "ยา 11" = 1,
                           R := "Stepper Motor ทำงาน สั่งconveyor เคลื่อที่ไปข้างหน้า" OR "ปุ่มClear",
                           PV := 1);
   "IEC_Counter_0_DB_37".CTUD(CU := ("Expected/Value_All".V = "Expected/Value_All".Expected_11) AND NOT "M11",
                           CD := "IEC_Counter_0_DB_1084".Q AND ("Barcode11" > 0) AND "ปุ่มยืนยันหน้า Screen",
                           PV := 5,
                           CV => "Barcode11");
   "M11" := "IEC_Counter_0_DB_37".QU;
   "IEC_Counter_0_DB_1085".CTU(CU := "ยา 12" = 1,
                           R := "Stepper Motor ทำงาน สั่งconveyor เคลื่อที่ไปข้างหน้า" OR "ปุ่มClear",
                           PV := 1);
   "IEC_Counter_0_DB_38".CTUD(CU := ("Expected/Value_All".V = "Expected/Value_All".Expected_12) AND NOT "M12",
                           CD := "IEC_Counter_0_DB_1085".Q AND ("Barcode12" > 0) AND "ปุ่มยืนยันหน้า Screen",
                           PV := 5,
                           CV => "Barcode12");
   "M12" := "IEC_Counter_0_DB_38".QU;
   "IEC_Counter_0_DB_1086".CTU(CU := "ยา 13" = 1,
                           R := "Stepper Motor ทำงาน สั่งconveyor เคลื่อที่ไปข้างหน้า" OR "ปุ่มClear",
                           PV := 1);
   "IEC_Counter_0_DB_39".CTUD(CU := ("Expected/Value_All".V = "Expected/Value_All".Expected_13) AND NOT "M13",
                           CD := "IEC_Counter_0_DB_1086".Q AND ("Barcode13" > 0) AND "ปุ่มยืนยันหน้า Screen",
                           PV := 5,
                           CV => "Barcode13");
   "M13" := "IEC_Counter_0_DB_39".QU;
   "IEC_Counter_0_DB_1087".CTU(CU := "ยา 14" = 1,
                           R := "Stepper Motor ทำงาน สั่งconveyor เคลื่อที่ไปข้างหน้า" OR "ปุ่มClear",
                           PV := 1);
   "IEC_Counter_0_DB_40".CTUD(CU := ("Expected/Value_All".V = "Expected/Value_All".Expected_14) AND NOT "M14",
                           CD := "IEC_Counter_0_DB_1087".Q AND ("Barcode14" > 0) AND "ปุ่มยืนยันหน้า Screen",
                           PV := 5,
                           CV => "Barcode14");
   "M14" := "IEC_Counter_0_DB_40".QU;
   "IEC_Counter_0_DB_1088".CTU(CU := "ยา 15" = 1,
                           R := "Stepper Motor ทำงาน สั่งconveyor เคลื่อที่ไปข้างหน้า" OR "ปุ่มClear",
                           PV := 1);
   "IEC_Counter_0_DB_41".CTUD(CU := ("Expected/Value_All".V = "Expected/Value_All".Expected_15) AND NOT "M15",
                           CD := "IEC_Counter_0_DB_1088".Q AND ("Barcode15" > 0) AND "ปุ่มยืนยันหน้า Screen",
                           PV := 5,
                           CV => "Barcode15");
   "M15" := "IEC_Counter_0_DB_41".QU;
   "IEC_Counter_0_DB_1089".CTU(CU := "ยา 16" = 1,
                           R := "Stepper Motor ทำงาน สั่งconveyor เคลื่อที่ไปข้างหน้า" OR "ปุ่มClear",
                           PV := 1);
   "IEC_Counter_0_DB_42".CTUD(CU := ("Expected/Value_All".V = "Expected/Value_All".Expected_16) AND NOT "M16",
                           CD := "IEC_Counter_0_DB_1089".Q AND ("Barcode16" > 0) AND "ปุ่มยืนยันหน้า Screen",
                           PV := 5,
                           CV => "Barcode16");
   "M16" := "IEC_Counter_0_DB_42".QU;
   "IEC_Counter_0_DB_1090".CTU(CU := "ยา 17" = 1,
                           R := "Stepper Motor ทำงาน สั่งconveyor เคลื่อที่ไปข้างหน้า" OR "ปุ่มClear",
                           PV := 1);
   "IEC_Counter_0_DB_43".CTUD(CU := ("Expected/Value_All".V = "Expected/Value_All".Expected_17) AND NOT "M17",
                           CD := "IEC_Counter_0_DB_1090".Q AND ("Barcode17" > 0) AND "ปุ่มยืนยันหน้า Screen",
                           PV := 5,
                           CV => "Barcode17");
   "M17" := "IEC_Counter_0_DB_43".QU;
   "IEC_Counter_0_DB_1091".CTU(CU := "ยา 18" = 1,
                           R := "Stepper Motor ทำงาน สั่งconveyor เคลื่อที่ไปข้างหน้า" OR "ปุ่มClear",
                           PV := 1);
   "IEC_Counter_0_DB_44".CTUD(CU := ("Expected/Value_All".V = "Expected/Value_All".Expected_18) AND NOT "M18",
                           CD := "IEC_Counter_0_DB_1091".Q AND ("Barcode18" > 0) AND "ปุ่มยืนยันหน้า Screen",
                           PV := 5,
                           CV => "Barcode18");
   "M18" := "IEC_Counter_0_DB_44".QU;
   "IEC_Counter_0_DB_1092".CTU(CU := "ยา 19" = 1,
                           R := "Stepper Motor ทำงาน สั่งconveyor เคลื่อที่ไปข้างหน้า" OR "ปุ่มClear",
                           PV := 1);
   "IEC_Counter_0_DB_45".CTUD(CU := ("Expected/Value_All".V = "Expected/Value_All".Expected_19) AND NOT "M19",
                           CD := "IEC_Counter_0_DB_1092".Q AND ("Barcode19" > 0) AND "ปุ่มยืนยันหน้า Screen",
                           PV := 5,
                           CV => "Barcode19");
   "M19" := "IEC_Counter_0_DB_45".QU;
   "IEC_Counter_0_DB_1093".CTU(CU := "ยา 20" = 1,
                           R := "Stepper Motor ทำงาน สั่งconveyor เคลื่อที่ไปข้างหน้า" OR "ปุ่มClear",
                           PV := 1);
   "IEC_Counter_0_DB_46".CTUD(CU := ("Expected/Value_All".V = "Expected/Value_All".Expected_20) AND NOT "M20",
                           CD := "IEC_Counter_0_DB_1093".Q AND ("Barcode20" > 0) AND "ปุ่มยืนยันหน้า Screen",
                           PV := 5,
                           CV => "Barcode20");
   "M20" := "IEC_Counter_0_DB_46".QU;
END_REGION

REGION Network 2
